(* IEC 61131-3 sources: daoli-st-library/DL_Device (part 6) *)

(* ---- FB_DL_SteamTrapMonitor.st ---- *)
(*==============================================================================
 * 组件名称 (Component)  : FB_DL_SteamTrapMonitor
 * 溯源说明 (Provenance): 道莅 clean-room 防御性实现（IEC 61131-3 纯净实现，闭源文档仅借语义，零代码行）
 * 所属子库 (Sublibrary) : DL_Device / Diagnostic
 * 当前版本 (Version)    : 1.0.0
 * 兼容性   (Platform)   : CODESYS 3.5 / TwinCAT 3 / 汇川 InoProShop / 施耐德
 *                         Machine Expert；纯 IEC 61131-3（第 3 版），仅用
 *                         Standard.library 的 TON / ABS / LIMIT / MAX
 * 组件分类 (Category)   : 功能块（FUNCTION_BLOCK）· 疏水阀堵塞/泄漏温差诊断
 * 功能一句话 (Summary)  : 用阀前/阀后温度差判断蒸汽疏水阀是正常、蒸汽泄漏（漏汽）
 *                         还是堵塞（不通），冷态停机时冻结全部故障判定。
 *
 * 本件存在的意义 (Why this unit exists)
 *   蒸汽系统节能诊断在全库零覆盖。疏水阀失效有两种相反形态：
 *   ① 漏汽（阀芯冲蚀常开）→ 阀后也被蒸汽烫热，温差变小，能耗与管网损失上升；
 *   ② 堵塞（阀芯卡死或结垢）→ 凝水积在阀前，阀前温度跌落，机组加热能力不足。
 *   两种都表现为「温差变小」，只能靠阀前温度是否达工况来区分——这就是本件
 *   判据的核心，也是它与普通温差异常报警的区别。
 *
 * 判据（公开工程判据，clean-room）
 *   正常   : fDelta >= fDeltaNormal
 *   漏汽   : fDelta <= fDeltaLeak 且 阀前温度达工况（fTin >= fTinMin）
 *   堵塞   : 阀前温度介于冷态带与工况下限之间（fTinMin × DL_COLD_RATIO <= fTin < fTinMin）
 *            且 fDelta <= fDeltaLeak
 *   冷态   : fTin < fTinMin × DL_COLD_RATIO → **工况未建立，冻结全部判定**（信息 0177）
 *   三条判据各带 tConfirm 持续确认窗，单拍越限不迁移（A5-D1 家族）。
 *   三条判据在数值上互斥（normal 要求 fDelta >= fDeltaNormal > fDeltaLeak；
 *   leak 要求 fTin >= fTinMin，blocked 要求 fTin < fTinMin），故不存在双判据
 *   同拍成立的两难情形——这是判据设计时就消除的，不靠优先级补丁。
 *
 * 冷态与堵塞的边界（规格冲突的落地方式，必须读）
 *   规格既要求「fTin < fTinMin 为工况未建立、冻结全部判定」，又要求「fTin < fTinMin
 *   （进出口均偏低、无温差）为堵塞」——同一条判据落两处。物理上二者靠「机组是否
 *   在跑」区分，本件引脚集没有机组运行信号，故用一条**相对冷态带**切分：
 *   fTinMin × DL_COLD_RATIO（0.5）以下视为停机冷态（冻结），该带与 fTinMin 之间
 *   视为「蒸汽已引入但被凝水淹没」= 堵塞特征。DL_COLD_RATIO 为件内经验常量，
 *   已在常量注释与偏离留档中声明；有运行信号的机型应把运行位并入 bEnable。
 *
 * 边界安全 (Boundary)
 *   ① fDeltaLeak >= fDeltaNormal（判据区间为空）或参数非有限 → 故障 0343、bValid = FALSE；
 *   ② 温度非有限 → 故障 0342，**保持上次判定与全部输出**（不迁移、不清状态）；
 *   ③ 冷态 → 信息 0177，冻结判定，健康投 eUnknown；
 *   ④ 落入正常带 → 信息 0176；
 *   ⑤ 健康映射集中在一处：漏汽 → eOutOfSpec（能耗越界）；堵塞 → eMaintenanceReq
 *      （需拆检）；故障 → eFailure；冷态/失能 → eUnknown；
 *   ⑥ CASE 落 ELSE 置 0344 并回 eFault；
 *   ⑦ 三条判据各用**独立 TON 实例**，绝不共用一只（R40）。
 *
 * 错误码    : 16#0003_0176 温差判据落入正常带——信息级，正常结论
 *             16#0003_0177 工况未建立（阀前温度低于冷态带），冻结判定——信息级，防误报
 *             16#0003_0342 温度输入非有限——故障级，保持上次判定
 *             16#0003_0343 判据阈值自相矛盾（fDeltaLeak >= fDeltaNormal）——故障级，bValid = FALSE
 *             16#0003_0344 状态机落 ELSE 兜底（非法状态）——故障级，回 eFault
 * 码位总账  : 16#0003_0176 用 / 16#0003_0177 用 ｜ 16#0003_0342 用 / 16#0003_0343 用 / 16#0003_0344 用
 * 状态机    : E_DL_TrapState（eIdle / eNormal / eLeak / eBlocked / eFault），CASE 含 ELSE 兜底，
 *             ELSE 置 16#0003_0344 并回 eFault；失能无条件回 eIdle
 * 采样约定  : 每任务周期调用一次；确认窗由 tConfirm 给定，不读系统时钟
 * 依赖说明  : 仅 Standard.library；健康出口引用 E_DL_Ne107Status（引用不重声明，R70③）
 * 验收向量  : V1 阀前 170 / 阀后 155（Δ15 >= 10）持续 30 s → eNormal，bNormal = TRUE，
 *                eErr = 0176，eHealth = eOk
 *             V2 阀前 165 / 阀后 162（Δ3、阀前达工况）持续 30 s → eLeak，bSteamLeak = TRUE，
 *                eHealth = eOutOfSpec
 *             V3 阀前 70 / 阀后 68（Δ2、介于冷态带 40 与 80 之间）持续 30 s → eBlocked，
 *                bBlocked = TRUE，eHealth = eMaintenanceReq（堵塞主向量）
 *             V4 阀前 30 / 阀后 28（低于冷态带 40）→ eIdle 冻结，eErr = 0177，eHealth = eUnknown
 *                （冷态防误报主向量）
 *             V5 fDeltaLeak = 12 > fDeltaNormal = 10 → 0343，bValid = FALSE，判据不成立
 *             V6 fTout = NaN → 0342，状态与输出保持上一拍（保持主向量）
 *             V7 温差在 9.9~10.1 抖动 → 单拍越限不迁移（确认窗主向量）
 * 红线自检  : 全局变量声明零使用 / 外部变量访问零使用 / 物理地址零使用 ｜ 纯 IEC 61131-3 ｜ 无除法
 *             浮点只用大小与容差比较 ｜ 无循环 ｜ 全变量双语同行注释 ｜ ENUM + CASE
 *             含 ELSE ｜ 三只 TON 在主体前部无条件刷新 ｜ 阈值常量化，无魔法数
 * 修订历史  : 2026-11-16  v1.0.0  首版入库（R22 · 批 3 · 设备诊断）
 *============================================================================*)

(*-----------------------------------------------------------------------------
 * 枚举: E_DL_TrapState（归属本功能块，同文件发布，全库唯一定义）
 * 含义: 疏水阀诊断相位。0 起步长 10。
 *-----------------------------------------------------------------------------*)
TYPE E_DL_TrapState :
(
    eIdle    := 0,     // 待机：未使能、冷态冻结或参数非法 / Idle, disabled, frozen cold state or illegal parameters
    eNormal  := 10,    // 正常：温差达到正常下限 / Normal, the temperature drop reaches the normal limit
    eLeak    := 20,    // 漏汽：温差过小且阀前已达工况 / Leaking, small drop with a live steam upstream
    eBlocked := 30,    // 堵塞：阀前温度跌落但蒸汽已引入 / Blocked, upstream cooled although steam was admitted
    eFault   := 99     // 故障：参数矛盾或非法状态 / Fault, contradictory parameters or an illegal state
);
END_TYPE

FUNCTION_BLOCK FB_DL_SteamTrapMonitor
VAR_INPUT
    fTin         : REAL;                       // 阀前温度 [degC] / upstream temperature [degC]
    fTout        : REAL;                       // 阀后温度 [degC] / downstream temperature [degC]
    fDeltaNormal : REAL := 10.0;               // 正常最小温差 [K]，须 > 0 / normal minimum temperature drop [K], must be > 0
    fDeltaLeak   : REAL := 5.0;                // 漏汽判定温差上限 [K]，须 >= 0 且 < fDeltaNormal / leak drop ceiling [K], below fDeltaNormal
    fTinMin      : REAL := 80.0;               // 蒸汽工况最低阀前温度 [degC]，须 > 0 / minimum live steam temperature [degC], must be > 0
    tConfirm     : TIME := T#30S;              // 判据确认时间 [ms] / criterion confirm time [ms]
    bEnable      : BOOL;                       // 使能 / enable
END_VAR
VAR_OUTPUT
    fDelta       : REAL;                       // 实测温差 = 阀前 − 阀后 [K] / measured temperature drop [K]
    bNormal      : BOOL;                       // 正常判定 / normal verdict
    bSteamLeak   : BOOL;                       // 漏汽判定 / steam leak verdict
    bBlocked     : BOOL;                       // 堵塞判定 / blocked verdict
    eHealth      : E_DL_Ne107Status;           // NE107 健康分级（引用唯一属主） / NE107 health status
    eErr         : UDINT;                      // 错误码，0 表示无错 / error code, 0 means no error
    bError       : BOOL;                       // 故障级标志，仅故障级错误置位 / fault-class flag, set only on fault-level codes
    bValid       : BOOL;                       // 输出可用标志 / outputs usable flag
END_VAR
VAR
    fbNormal     : TON;                        // 正常判据确认窗，段 7 无条件刷新 [ms] / normal criterion confirm window
    fbLeak       : TON;                        // 漏汽判据确认窗，段 7 无条件刷新 [ms] / leak criterion confirm window
    fbBlocked    : TON;                        // 堵塞判据确认窗，段 7 无条件刷新 [ms] / blocked criterion confirm window
    _eState      : E_DL_TrapState := E_DL_TrapState.eIdle; // 当前相位 / current phase
    _bInit       : BOOL := FALSE;              // 首扫标志，初值 FALSE 取非判定 / first-scan flag, tested negated
    _bParamBad   : BOOL;                       // 参数非法标志 / illegal parameter flag
    _bFiniteBad  : BOOL;                       // 输入非有限标志 / non-finite input flag
    _bIllegal    : BOOL;                       // 非法状态标志 / illegal state flag
    _bCold       : BOOL;                       // 冷态（工况未建立）标志 / cold state, the operating condition is not established
    _bCondNormal : BOOL;                       // 正常判据条件 / normal criterion condition
    _bCondLeak   : BOOL;                       // 漏汽判据条件 / leak criterion condition
    _bCondBlock  : BOOL;                       // 堵塞判据条件 / blocked criterion condition
    _bBrkNormal  : BOOL;                       // 正常确认计时器断输入一拍 / normal timer one-scan break
    _bBrkLeak    : BOOL;                       // 漏汽确认计时器断输入一拍 / leak timer one-scan break
    _bBrkBlock   : BOOL;                       // 堵塞确认计时器断输入一拍 / blocked timer one-scan break
    _tConfirmUse : TIME := T#30S;              // 生效确认时间 [ms]，已钳位 / effective confirm time, clamped
    _fDeltaHeld  : REAL;                       // 温差保持量 [K] / held temperature drop [K]
    _fColdLimit  : REAL := 40.0;               // 冷态带上限 [degC] = fTinMin × 冷态比 / cold band ceiling
END_VAR
VAR CONSTANT
    DL_VAL_LIM     : REAL := 1.0E6;            // 有限性判定的绝对值上限 [degC] / finiteness ceiling [degC]
    DL_DELTA_N_MN  : REAL := 0.0;              // 正常温差下限 [K]，须严格大于 / normal drop floor, strictly greater
    DL_DELTA_L_MN  : REAL := 0.0;              // 漏汽温差下限 [K] / leak drop floor [K]
    DL_TIN_MIN_MN  : REAL := 0.0;              // 工况温度下限 [degC]，须严格大于 / live steam temperature floor, strictly greater
    DL_COLD_RATIO  : REAL := 0.5;              // 冷态带相对工况下限的比例 [倍]，件内经验值 / cold band ratio, an empirical in-unit value
    DL_DELTA_MAX   : REAL := 1000.0;           // 温差合理上限 [K]，仅用于出口钳位 / sane drop ceiling [K], outlet clamping only
    DL_CONF_MAX_MS : DINT := 3600000;          // 确认时间上限 [ms]，一小时 / confirm time ceiling, one hour
    DL_TIME_ZERO   : TIME := T#0MS;            // 时间零值基准 [ms] / time zero reference
    DL_EPS         : REAL := 1.0E-6;           // 浮点比较容差 [K] / float comparison tolerance [K]
END_VAR

(*------------------------------------------------------------------------------
 * 段 1｜每拍预置（判定输出与保持量在段 9 单点写入）
 *      Per-scan presets, the verdicts are written only in segment nine
 *-----------------------------------------------------------------------------*)
eErr         := 16#0000_0000;                  // 错误码每拍重算 / error code recomputed every scan
bError       := FALSE;                         // 故障标志每拍重算 / fault flag recomputed every scan
bValid       := FALSE;                         // 可用标志每拍重算 / usable flag recomputed every scan
bNormal      := FALSE;                         // 正常判定每拍重算 / normal verdict recomputed
bSteamLeak   := FALSE;                         // 漏汽判定每拍重算 / leak verdict recomputed
bBlocked     := FALSE;                         // 堵塞判定每拍重算 / blocked verdict recomputed
_bParamBad   := FALSE;                         // 参数非法标志预清零 / parameter flag pre-cleared
_bFiniteBad  := FALSE;                         // 非有限标志预清零 / non-finite flag pre-cleared
_bIllegal    := FALSE;                         // 非法状态标志预清零 / illegal state flag pre-cleared
_bCold       := FALSE;                         // 冷态标志预清零 / cold flag pre-cleared
_bCondNormal := FALSE;                         // 正常条件预置 FALSE / normal condition preset FALSE
_bCondLeak   := FALSE;                         // 漏汽条件预置 FALSE / leak condition preset FALSE
_bCondBlock  := FALSE;                         // 堵塞条件预置 FALSE / blocked condition preset FALSE

(*------------------------------------------------------------------------------
 * 段 2｜首扫初始化（判定从待机起，不继承任何历史结论）
 *      First-scan initialisation, no historical verdict is inherited
 *-----------------------------------------------------------------------------*)
IF NOT _bInit THEN
    _eState     := E_DL_TrapState.eIdle;       // 相位待机 / phase idle
    _fDeltaHeld := 0.0;                        // 温差保持量 0 [K] / held drop zero
    _bBrkNormal := TRUE;                       // 正常确认窗从零开始 / normal window starts from zero
    _bBrkLeak   := TRUE;                       // 漏汽确认窗从零开始 / leak window starts from zero
    _bBrkBlock  := TRUE;                       // 堵塞确认窗从零开始 / blocked window starts from zero
    _bInit      := TRUE;                       // 首扫只做一次 / the first scan runs once
END_IF

(*------------------------------------------------------------------------------
 * 段 3｜参数闸门（判据区间必须非空，否则判据无意义）
 *      Parameter gate, the criteria intervals must not be empty
 *-----------------------------------------------------------------------------*)
IF (fDeltaNormal <> fDeltaNormal) OR (ABS(fDeltaNormal) > DL_VAL_LIM) OR (fDeltaNormal <= DL_DELTA_N_MN) THEN
    _bParamBad := TRUE;                        // 正常温差非法 / normal drop illegal
END_IF
IF (fDeltaLeak <> fDeltaLeak) OR (ABS(fDeltaLeak) > DL_VAL_LIM) OR (fDeltaLeak < DL_DELTA_L_MN) THEN
    _bParamBad := TRUE;                        // 漏汽温差非法 / leak drop illegal
END_IF
IF (fDeltaLeak >= fDeltaNormal) OR ((fDeltaNormal - fDeltaLeak) <= DL_EPS) THEN
    _bParamBad := TRUE;                        // 区间为空：判据自相矛盾 / empty interval, contradictory criteria
END_IF
IF (fTinMin <> fTinMin) OR (ABS(fTinMin) > DL_VAL_LIM) OR (fTinMin <= DL_TIN_MIN_MN) THEN
    _bParamBad := TRUE;                        // 工况温度非法 / live steam temperature illegal
END_IF

(*------------------------------------------------------------------------------
 * 段 4｜温度有限性（区间判据同时拦 NaN 与 ±Inf）
 *      Temperature finiteness, the interval test catches NaN and infinity
 *-----------------------------------------------------------------------------*)
IF (fTin < -DL_VAL_LIM) OR (fTin > DL_VAL_LIM) THEN
    _bFiniteBad := TRUE;                       // 阀前温度非有限 / upstream temperature non-finite
END_IF
IF (fTout < -DL_VAL_LIM) OR (fTout > DL_VAL_LIM) THEN
    _bFiniteBad := TRUE;                       // 阀后温度非有限 / downstream temperature non-finite
END_IF

(*------------------------------------------------------------------------------
 * 段 5｜温差与冷态带（冷态带由工况下限按比例导出，件内常量）
 *      Temperature drop and the cold band derived from the live steam limit
 *-----------------------------------------------------------------------------*)
IF NOT _bFiniteBad THEN
    _fDeltaHeld := fTin - fTout;               // 实测温差 [K] / measured drop
    _fColdLimit := fTinMin * DL_COLD_RATIO;    // 冷态带上限 [degC] / cold band ceiling
    _bCold      := (fTin < _fColdLimit);       // 冷态判据：明显停机 / cold test, clearly shut down
END_IF

(*------------------------------------------------------------------------------
 * 段 6｜三条判据条件（数值上互斥：由阈值关系结构性保证，不靠优先级补丁）
 *      The three criteria are mutually exclusive by construction
 *-----------------------------------------------------------------------------*)
IF (NOT _bFiniteBad) AND (NOT _bParamBad) THEN
    _bCondNormal := (_fDeltaHeld >= fDeltaNormal);                       // 正常：温差达正常下限
    _bCondLeak   := (_fDeltaHeld <= fDeltaLeak) AND (fTin >= fTinMin);   // 漏汽：温差小且阀前已达工况
    _bCondBlock  := (_fDeltaHeld <= fDeltaLeak) AND (fTin >= _fColdLimit) AND (fTin < fTinMin); // 堵塞：蒸汽已引入但阀前跌落
END_IF

(*------------------------------------------------------------------------------
 * 段 7｜三只确认计时器无条件刷新（R40：CASE 之外每拍必调，各判据各一只）
 *      Three confirm timers refreshed unconditionally, one instance per criterion
 *-----------------------------------------------------------------------------*)
_tConfirmUse := tConfirm;                      // 确认时间直取引脚 [ms] / confirm time from the pin
IF TIME_TO_DINT(_tConfirmUse) > DL_CONF_MAX_MS THEN
    _tConfirmUse := DINT_TO_TIME(DL_CONF_MAX_MS); // 超上限钳位（无专用码位，R90 不新开码） / clamped
END_IF
IF TIME_TO_DINT(_tConfirmUse) < 0 THEN
    _tConfirmUse := DL_TIME_ZERO;              // 负时间结构性不可达，兜底为 0 / structurally unreachable fallback
END_IF

fbNormal(IN := _bCondNormal AND bEnable AND (NOT _bBrkNormal), PT := _tConfirmUse); // 正常确认窗
_bBrkNormal := FALSE;                          // 断输入拍在调用后自清 / break self-cleared after the call

fbLeak(IN := _bCondLeak AND bEnable AND (NOT _bBrkLeak), PT := _tConfirmUse); // 漏汽确认窗
_bBrkLeak := FALSE;                            // 断输入拍在调用后自清 / break self-cleared

fbBlocked(IN := _bCondBlock AND bEnable AND (NOT _bBrkBlock), PT := _tConfirmUse); // 堵塞确认窗
_bBrkBlock := FALSE;                           // 断输入拍在调用后自清 / break self-cleared

(*------------------------------------------------------------------------------
 * 段 8｜相位机（非有限拍整段跳过：保持上次判定，②）
 *      Phase machine, skipped entirely on a non-finite scan to hold the last verdict
 *-----------------------------------------------------------------------------*)
IF NOT _bFiniteBad THEN
    (* 温度坏值拍整段跳过：不迁移、不清结论，保持上次判定（②），仅由码位链报 0342 *)
    (* A non-finite scan skips the whole block, the last verdict is held *)
    IF _bParamBad THEN
        _eState := E_DL_TrapState.eFault;      // 判据自相矛盾：转故障 / contradictory criteria go to fault
    ELSIF NOT bEnable THEN
        _eState := E_DL_TrapState.eIdle;       // 失能回待机 / disabled, back to idle
        _bBrkNormal := TRUE;                   // 三只确认窗全部重启 / every window restarts
        _bBrkLeak   := TRUE;                   // 漏汽窗重启 / leak window restarts
        _bBrkBlock  := TRUE;                   // 堵塞窗重启 / blocked window restarts
    ELSE
        CASE _eState OF

            E_DL_TrapState.eIdle:                  // 待机：冷态冻结，工况建立后按判据进入
                IF _bCold THEN
                    _eState := E_DL_TrapState.eIdle; // 工况未建立，冻结（0177 在段 10） / condition not established, frozen
                ELSIF fbNormal.Q THEN
                    _eState := E_DL_TrapState.eNormal; // 进正常相 / enter normal
                ELSIF fbLeak.Q THEN
                    _eState := E_DL_TrapState.eLeak;   // 进漏汽相 / enter leak
                ELSIF fbBlocked.Q THEN
                    _eState := E_DL_TrapState.eBlocked; // 进堵塞相 / enter blocked
                END_IF

            E_DL_TrapState.eNormal:                // 正常：判据迁移
                IF _bCold THEN
                    _eState := E_DL_TrapState.eIdle;   // 工况消失，回冻结 / the condition is lost, freeze
                ELSIF fbLeak.Q THEN
                    _eState := E_DL_TrapState.eLeak;   // 转漏汽 / switch to leak
                ELSIF fbBlocked.Q THEN
                    _eState := E_DL_TrapState.eBlocked; // 转堵塞 / switch to blocked
                END_IF

            E_DL_TrapState.eLeak:                  // 漏汽：判据迁移
                IF _bCold THEN
                    _eState := E_DL_TrapState.eIdle;   // 工况消失，回冻结 / freeze again
                ELSIF fbNormal.Q THEN
                    _eState := E_DL_TrapState.eNormal; // 恢复正常 / back to normal
                ELSIF fbBlocked.Q THEN
                    _eState := E_DL_TrapState.eBlocked; // 转堵塞 / switch to blocked
                END_IF

            E_DL_TrapState.eBlocked:               // 堵塞：判据迁移
                IF _bCold THEN
                    _eState := E_DL_TrapState.eIdle;   // 工况消失（彻底冷机），回冻结 / freeze again
                ELSIF fbNormal.Q THEN
                    _eState := E_DL_TrapState.eNormal; // 恢复正常 / back to normal
                ELSIF fbLeak.Q THEN
                    _eState := E_DL_TrapState.eLeak;   // 转漏汽 / switch to leak
                END_IF

            E_DL_TrapState.eFault:                 // 故障：参数恢复即回待机
                IF (NOT _bParamBad) AND (NOT _bFiniteBad) THEN
                    _eState := E_DL_TrapState.eIdle;   // 原因消失 / the cause is gone
                END_IF

            ELSE
                _bIllegal := TRUE;                 // 标记非法状态 / flag the illegal state
                _eState   := E_DL_TrapState.eFault; // 回故障态 / back to the fault state
        END_CASE
    END_IF
END_IF

(*------------------------------------------------------------------------------
 * 段 9｜出口单点写入（判定与温差唯一写入点）
 *      Single write point of the verdicts and the temperature drop
 *-----------------------------------------------------------------------------*)
fDelta := LIMIT(-DL_DELTA_MAX, _fDeltaHeld, DL_DELTA_MAX); // 温差出口钳进合理域 [K] / the drop is clamped
bNormal    := (_eState = E_DL_TrapState.eNormal);   // 正常判定出口 / normal verdict outlet
bSteamLeak := (_eState = E_DL_TrapState.eLeak);     // 漏汽判定出口 / leak verdict outlet
bBlocked   := (_eState = E_DL_TrapState.eBlocked);  // 堵塞判定出口 / blocked verdict outlet

(*------------------------------------------------------------------------------
 * 段 10｜码位优先级链与健康分级（映射集中在此，不散落实现体）
 *      Code priority chain and health grading, the mapping lives in one place
 *-----------------------------------------------------------------------------*)
IF _bIllegal THEN
    eErr   := 16#0003_0344;                    // 故障级：状态机兜底 / fault: state machine fallback
    bError := TRUE;                            // 置故障标志 / raise the fault flag
ELSIF _bParamBad THEN
    eErr   := 16#0003_0343;                    // 故障级：判据阈值自相矛盾 / fault: contradictory thresholds
    bError := TRUE;                            // 置故障标志 / raise the fault flag
ELSIF _bFiniteBad THEN
    eErr   := 16#0003_0342;                    // 故障级：温度输入非有限 / fault: non-finite temperature
    bError := TRUE;                            // 置故障标志 / raise the fault flag
ELSIF _bCold THEN
    eErr   := 16#0003_0177;                    // 信息级：工况未建立，冻结判定 / informational: condition not established
ELSIF _eState = E_DL_TrapState.eNormal THEN
    eErr   := 16#0003_0176;                    // 信息级：判据落入正常带 / informational: inside the normal band
END_IF

IF _bParamBad OR _bFiniteBad OR _bIllegal THEN
    eHealth := E_DL_Ne107Status.eFailure;      // 无判定能力：失效 / no verdict capability
ELSIF _eState = E_DL_TrapState.eLeak THEN
    eHealth := E_DL_Ne107Status.eOutOfSpec;    // 漏汽：能耗与管网越界，仍可运行 / leaking, out of specification
ELSIF _eState = E_DL_TrapState.eBlocked THEN
    eHealth := E_DL_Ne107Status.eMaintenanceReq; // 堵塞：需拆检 / blocked, maintenance required
ELSIF (_eState = E_DL_TrapState.eNormal) AND bEnable THEN
    eHealth := E_DL_Ne107Status.eOk;           // 正常 / normal
ELSE
    eHealth := E_DL_Ne107Status.eUnknown;      // 冷态或失能：无结论 / cold or disabled, no verdict
END_IF

IF bError THEN
    bValid := FALSE;                           // 故障级：输出不可用 / fault: outputs unusable
ELSIF _bCold THEN
    bValid := FALSE;                           // 冷态：判定被冻结，输出不可用 / cold: the verdict is frozen
ELSIF NOT bEnable THEN
    bValid := FALSE;                           // 失能：输出不可用 / disabled: unusable
ELSE
    bValid := TRUE;                            // 判定可用 / verdict usable
END_IF

END_FUNCTION_BLOCK

(* ---- FB_DL_StrainThermalCreepAdaptive.st ---- *)
(*
    FB_DL_StrainThermalCreepAdaptive —— 应变桥温漂与蠕变自适应补偿（含空载窗口自动重学零点）
    ------------------------------------------------------------------
    组件名    : FB_DL_StrainThermalCreepAdaptive
    分类      : DL_Device / Weighing Compensation（称重与测力补偿）
    一句话功能: 在线扣除应变桥的温漂与载荷蠕变，并在空载窗口自动重学零点，
                同时用「载荷是否真为空」判据防止把真实载荷学成漂移。
    复杂度    : C3
    版本      : v1.0.0
    开源溯源  : 无（clean-room 自研，未借鉴任何开源实现）
    平台      : 纯 IEC 61131-3（TON / R_TRIG / ABS / TIME_TO_REAL 标准转换），目标编译器
                RuSTy 1.0.8，兼容 CODESYS 3.5 / TwinCAT 3 / 汇川 InoProShop / Machine Expert；
                无 PROPERTY、无 VLA、无 FOR..DOWNTO、无 AS 类方言
    ------------------------------------------------------------------
    功能说明  : ① 温漂：fTempCorrMv = fTempCoefMvPerC × (fTempC − fRefTempC)，从原始桥压减掉；
                ② 零点：fCorrected = fRawMv − fTempCorrMv − fZeroMv，零点由空载学习维护；
                ③ 蠕变：fCreepCorrMv = fCorrected × fCreepCoefPctPerMin × 0.01 × tHoldMin，
                   方向随 fCorrected 的符号自动跟随载荷方向（负载荷得到负补偿量）；
                ④ 空载学习：bNoLoadWindow = TRUE 且持续 ≥ tLearnMinMs（TON 无条件刷新）→ 进
                   eLearn，用一阶低通（系数固定 0.05，见代理假设）把「温漂修正后、零点修正前」
                   的值学成新零点；窗口消失立即退出并冻结零点；
                ⑤ 防误学：学习期间若 |温漂修正后值| 超 fNoLoadMaxMv（载荷比 > 1）→ 判「并非空载」，
                   退出 eLearn 回 eRun 并置 bLearnRejected 单拍位；同一空载窗口内不再重试
                   （_bRejLatch 在窗口消失时清除），避免窗口内反复进出打摆；
                ⑥ 温度或原始值非有限 → eFault，且 fOutMv 保持上一次有效值（保持而非清零）。
    量纲链    : fTempCoefMvPerC [mV/°C] × (fTempC − fRefTempC) [°C] → fTempCorrMv [mV]（°C 约去）；
                fRawMv [mV] − fTempCorrMv [mV] → _fRawTemp [mV]（零点修正前）；
                _fRawTemp [mV] − fZeroMv [mV] → fCorrected [mV]（零点修正后）；
                fCorrected [mV] × fCreepCoefPctPerMin [%/min] × 0.01 [1/%] × tHoldMin [min]
                    → fCreepCorrMv [mV]（%/min × min = %，× 0.01 无因次，只剩 mV）；
                fOutMv = fCorrected [mV] − fCreepCorrMv [mV] → [mV]；
                _fLoadRatio = |_fRawTemp| [mV] ÷ _fNoLoadGuard [mV] → [-]（判载荷比与 1.0 直比）。
                全程无「温度与毫伏相加」「时间与毫伏相加」，量纲链逐段闭合。
    代理假设  : （R95 三句声明）① 代理值 = 低通系数固定 0.05，隐含标称扫描周期 10 ms，
                对应零点学习时间常数 τ ≈ 0.2 s；② 覆盖范围 = 5 ms ~ 20 ms 的周期任务
                （时间常数随之在 0.1 s ~ 0.4 s 间变化，只影响学习快慢，不影响零点收敛方向）；
                ③ 覆盖不到的区间（< 2 ms 或 > 50 ms 的任务）由现场加长 tLearnMinMs 与空载窗口
                驻留时长补偿，本件不提供自适应系数。
    交付门槛  : 本件使用 TIME_TO_REAL 标准转换做承载时长换算，须在 CODESYS / TwinCAT /
                InoProShop 三平台各编译验证一次（R64）。
    状态机    : eInit(0) --使能且输入有限且组态合法--> eRun(10)
                eRun --空载窗口持续到（tonLearn.Q）且本窗口未拒学过--> eLearn(20)
                eLearn --窗口消失--> eRun（零点冻结）；--载荷比 > 1--> eRun（拒学 + 单拍位）
                eRun/eLearn --失能--> eHold(30)（冻结保持末次有效输出与累计）
                eHold --重新使能--> eRun
                任意相 --输入非有限或组态非法--> eFault(90)
                eFault 的唯一解除路径 = bReset 上升沿（见段 8 与复位作用域声明）
    失能语义  : bEnable = FALSE → eHold，fOutMv 冻结保持末次有效值，蠕变累计与零点学习全部冻结
                （取「冻结保持」而非「降级清零」：称重输出清零会被上位当作零载荷，属伪造计量事实）。
    复位作用域: bReset 上升沿①清 _bFaultLatch / _bBadIn / _bCfgBad；②清 _fZero 与
                _fHoldBaseMin（零点与承载累计一并归零，须重新学习）；③清 _bRejLatch；
                ④迁相回 eInit；⑤不清 _fOutHold（补偿输出不因复位跳变），_bHoldValid 保留。
    防御口径  : NaN 用自反 f<>f；±Inf 用 (f−f)<>(f−f)；另设幅值域闸 ABS(f) > 1.0E30。
                除子三类：DL_ST_MS_PER_MIN = 60000.0 与 DL_ST_PCT_TO_RATIO = 0.01 为具名常量，
                结构上不可能为零；载荷比除子 _fNoLoadGuard 由 fNoLoadMaxMv 经两级下限兜底后
                才参与除法（R117 两级回退）。
                计算结果写入保持槽 _fOutHold 之前必须过非有限闸（R133），污染数据不进保持槽。
    规格偏离  : 派单把学习最短时长写作 fLearnMinMs，其实际类型为 TIME；本库规范 1.2 规定
                时间量前缀为 t，故落为 tLearnMinMs，语义不变。按 R190 归因唯一补充
                bCfgErr / bDataErr 两个诊断位，使两条故障成因各自可观测。
    码位说明  : 本件按零码位范式交付，不分配 16# 事件码；学习结果与故障一律经
                eState / bLearnRejected / bFaultOut / bCfgErr / bDataErr 组合观测。
    修订记录  : 2026-11-24 v1.0.0 首次入库（R87 批 · #3）
*)
TYPE E_DL_StrainCompState :
(
    eInit   := 0,     // 初始化：首扫或复位后，尚无可信输出 | init, no trustworthy output yet
    eRun    := 10,    // 运行：温漂 + 零点 + 蠕变三项全补偿 | running, thermal, zero and creep all compensated
    eLearn  := 20,    // 学习：空载窗口内低通重学零点，蠕变累计冻结 | learning the zero in a no-load window
    eHold   := 30,    // 保持：失能冻结末次有效输出与累计 | hold, disabled, last valid output frozen
    eFault  := 90     // 故障：输入非有限或组态非法，锁存至复位沿 | fault latched until the reset edge
);
END_TYPE

FUNCTION_BLOCK FB_DL_StrainThermalCreepAdaptive
VAR_INPUT
    bEnable             : BOOL;                   // 使能电平，TRUE = 允许补偿与学习 | enable level, TRUE = compensation and learning
    bReset              : BOOL;                   // 复位请求，上升沿生效 | reset request, rising-edge active
    fRawMv              : REAL;                   // 应变桥原始输出 [mV] | raw bridge output [mV]
    fTempC              : REAL;                   // 桥体温度 [°C] | bridge temperature [degC]
    fRefTempC           : REAL := 20.0;           // 参考温度（补偿零点温度）[°C] | reference temperature [degC]
    fTempCoefMvPerC     : REAL := 0.0;            // 温度系数 [mV/°C]，正负均合法 | temperature coefficient [mV/degC]
    fCreepCoefPctPerMin : REAL := 0.0;            // 蠕变系数 [%/min]，须非负 | creep coefficient [%/min], non-negative
    bNoLoadWindow       : BOOL;                   // 空载窗口（上位给出：工位确认为空载）| no-load window from the supervisor
    tLearnMinMs         : TIME := T#2S;           // 空载最短驻留时长，达到才允许学习 [ms] | minimum no-load dwell [ms]
    fNoLoadMaxMv        : REAL := 0.5;            // 空载带半宽，超出即判非空载 [mV] | no-load band half width [mV]
END_VAR
VAR_OUTPUT
    eState              : E_DL_StrainCompState;          // 主状态，供 HMI 使用 | main state for HMI
    fOutMv              : REAL;                   // 补偿后输出（去皮净载荷）[mV] | compensated output [mV]
    fTempCorrMv         : REAL;                   // 本拍温漂补偿量 [mV] | thermal correction this scan [mV]
    fCreepCorrMv        : REAL;                   // 本拍蠕变补偿量 [mV] | creep correction this scan [mV]
    fZeroMv             : REAL;                   // 当前生效零点 [mV] | active zero offset [mV]
    bLearnRejected      : BOOL;                   // 学习被拒事件位，单拍 | learning rejection event, single scan
    bFaultOut           : BOOL;                   // 故障汇总位 | fault aggregate
    bCfgErr             : BOOL;                   // 组态非法诊断位（归因唯一，R190）| bad-configuration flag
    bDataErr            : BOOL;                   // 数据非有限诊断位（归因唯一，R190）| non-finite data flag
END_VAR
VAR
    rtReset             : R_TRIG;                 // 复位上升沿实例，每拍无条件刷新 | reset rising-edge instance
    tonHold             : TON;                    // 承载时长分片计时，自复位，每拍无条件刷新 | load-hold slice timer, self-resetting
    tonLearn            : TON;                    // 空载窗口驻留计时，每拍无条件刷新 | no-load dwell timer
    _eState             : E_DL_StrainCompState := E_DL_StrainCompState.eInit; // 状态机内部当前态 | internal current state
    _bInit              : BOOL := TRUE;           // 首扫初始化标志，含零点与累计状态 | first-scan init flag
    _bResetLatch        : BOOL := FALSE;          // 复位沿锁存量，本拍末清除 | reset-edge latch, cleared at scan end
    _bFaultLatch        : BOOL := FALSE;          // 故障锁存位 | fault latch
    _bBadIn             : BOOL := FALSE;          // 输入非有限成因位 | non-finite input cause
    _bCfgBad            : BOOL := FALSE;          // 组态非法成因位 | bad configuration cause
    _bRejLatch          : BOOL := FALSE;          // 拒学锁存，空载窗口消失时清除 | rejection latch, cleared when the window drops
    _bHoldValid         : BOOL := FALSE;          // 保持槽已有有效值标志 | holder contains a valid value
    _bLoadNow           : BOOL := FALSE;          // 本拍存在载荷（超空载带）| load present this scan
    _fZero              : REAL := 0.0;            // 学习得到的零点 [mV] | learned zero offset [mV]
    _fTempCorr          : REAL := 0.0;            // 温漂补偿量 [mV] | thermal correction [mV]
    _fRawTemp           : REAL := 0.0;            // 温漂修正后、零点修正前的值 [mV] | thermally corrected, pre-zero [mV]
    _fCorrected         : REAL := 0.0;            // 温漂与零点均修正后的值 [mV] | fully corrected value [mV]
    _fCreepCorr         : REAL := 0.0;            // 蠕变补偿量 [mV] | creep correction [mV]
    _fOut               : REAL := 0.0;            // 本拍补偿输出 [mV] | compensated output this scan [mV]
    _fOutHold           : REAL := 0.0;            // 输出保持槽，只写已过非有限闸的值 [mV] | output holder, gated before writing [mV]
    _fNoLoadGuard       : REAL := 0.0;            // 空载带半宽的兜底值 [mV]，作除法除子 | no-load band with floor, used as divisor [mV]
    _fLoadRatio         : REAL := 0.0;            // 载荷比 [-] = |值| ÷ 空载带半宽 | load ratio, dimensionless
    _fHoldBaseMin       : REAL := 0.0;            // 已满片承载时长基值 [min] | accumulated whole-slice hold time [min]
    _fHoldMin           : REAL := 0.0;            // 参与蠕变计算的承载时长 [min] | hold time used by the creep model [min]
END_VAR
VAR CONSTANT
    DL_ST_EPS           : REAL := 1.0E-6;         // 浮点判零容差 [mV] | float zero tolerance [mV]
    DL_ST_MAG_MAX       : REAL := 1.0E30;         // 有限幅值域闸上限 [mV] | magnitude domain bound [mV]
    DL_ST_BAND_FLOOR    : REAL := 1.0E-3;         // 空载带半宽下限兜底 [mV] | no-load band floor [mV]
    DL_ST_LPF_ALPHA     : REAL := 0.05;           // 零点学习低通系数 [-]，见代理假设三句 | zero-learning low-pass coefficient
    DL_ST_MS_PER_MIN    : REAL := 60000.0;        // 毫秒与分钟换算常量 [ms/min] | milliseconds per minute
    DL_ST_PCT_TO_RATIO  : REAL := 0.01;           // 百分数转无因次常量 [1/%] | percent to ratio constant
    DL_ST_SLICE_MIN     : REAL := 60.0;           // 承载时长分片宽度 [min]（对应 TON 的 1 h 量程）| hold slice width [min]
    DL_ST_HOLD_MAX_MIN  : REAL := 1000000.0;      // 承载时长基值饱和上限 [min]，防浮点溢出 | hold-time saturation bound [min]
END_VAR

METHOD ClampToBand : REAL
(*
    把补偿量钳到 ±带宽，防止系数误配时补偿量把输出打穿。纯函数，无跨拍状态。
    Clamp a correction to a symmetric band so a mis-parameterised coefficient cannot saturate the output.
*)
VAR_INPUT
    fIn   : REAL;                                 // 待钳补偿量 [mV] | correction to clamp [mV]
    fBand : REAL;                                 // 对称带宽（已兜底为正）[mV] | symmetric band, floored positive [mV]
END_VAR
ClampToBand := fIn;                               // 直通后按两侧硬界饱和 | straight-through, saturated below
IF ClampToBand > fBand THEN
    ClampToBand := fBand;                         // 正向钳到 +带宽 [mV] | clamp to the positive band
END_IF
IF ClampToBand < (0.0 - fBand) THEN
    ClampToBand := 0.0 - fBand;                   // 负向钳到 −带宽 [mV] | clamp to the negative band
END_IF
END_METHOD

// 段 1｜输出预置与首扫初始化（含零点与累计状态，故必须有 _bInit，R310）
// segment 1, output presets and first-scan initialisation; the zero and accumulators require _bInit
fTempCorrMv := 0.0;                                // 预置温漂补偿 0 [mV] | preset zero thermal correction [mV]
fCreepCorrMv := 0.0;                               // 预置蠕变补偿 0 [mV] | preset zero creep correction [mV]
bLearnRejected := FALSE;                           // 预置无拒学事件（清零归属本段，R256）| preset no rejection event
_bBadIn := FALSE;                                  // 预置输入有限 | preset finite input
_bCfgBad := FALSE;                                 // 预置组态合法 | preset legal configuration
_bLoadNow := FALSE;                                // 预置无载荷 | preset no load
IF _bInit THEN
    _bInit := FALSE;                               // 首扫只执行一次 | runs once on the first scan
    _eState := E_DL_StrainCompState.eInit;                // 首扫状态回初相 | initialise the state
    _fZero := 0.0;                                 // 首扫零点归零 [mV]，由空载学习建立 | initial zero [mV]
    _fHoldBaseMin := 0.0;                          // 首扫承载时长归零 [min] | initial hold time [min]
    _fHoldMin := 0.0;                              // 首扫参与量归零 [min] | initial hold time for the model [min]
    _bRejLatch := FALSE;                           // 首扫清拒学锁存 | clear the rejection latch
    _bHoldValid := FALSE;                          // 首扫无有效保持值 | no valid holder value yet
END_IF

// 段 2｜非有限闸：NaN 自反 + Inf 自减 + 幅值域，逐个浮点入参枚举（R4 / R151 / R272）
// segment 2, non-finite gate over every REAL input: NaN self-reflexive, Inf by self-subtraction, magnitude bound
IF (fRawMv <> fRawMv) OR ((fRawMv - fRawMv) <> (fRawMv - fRawMv)) THEN
    _bBadIn := TRUE;                               // 原始桥压 NaN 或 ±Inf | raw bridge output NaN or infinity
END_IF
IF ABS(fRawMv) > DL_ST_MAG_MAX THEN
    _bBadIn := TRUE;                               // 原始桥压超幅值域 | raw bridge output beyond the magnitude domain
END_IF
IF (fTempC <> fTempC) OR ((fTempC - fTempC) <> (fTempC - fTempC)) THEN
    _bBadIn := TRUE;                               // 温度 NaN 或 ±Inf | temperature NaN or infinity
END_IF
IF ABS(fTempC) > DL_ST_MAG_MAX THEN
    _bBadIn := TRUE;                               // 温度超幅值域 | temperature beyond the magnitude domain
END_IF
IF (fRefTempC <> fRefTempC) OR ((fRefTempC - fRefTempC) <> (fRefTempC - fRefTempC)) THEN
    _bBadIn := TRUE;                               // 参考温度 NaN 或 ±Inf | reference temperature NaN or infinity
END_IF
IF ABS(fRefTempC) > DL_ST_MAG_MAX THEN
    _bBadIn := TRUE;                               // 参考温度超幅值域 | reference temperature beyond the magnitude domain
END_IF
IF (fTempCoefMvPerC <> fTempCoefMvPerC) OR ((fTempCoefMvPerC - fTempCoefMvPerC) <> (fTempCoefMvPerC - fTempCoefMvPerC)) THEN
    _bBadIn := TRUE;                               // 温度系数 NaN 或 ±Inf | temperature coefficient NaN or infinity
END_IF
IF ABS(fTempCoefMvPerC) > DL_ST_MAG_MAX THEN
    _bBadIn := TRUE;                               // 温度系数超幅值域 | temperature coefficient beyond the magnitude domain
END_IF
IF (fCreepCoefPctPerMin <> fCreepCoefPctPerMin) OR ((fCreepCoefPctPerMin - fCreepCoefPctPerMin) <> (fCreepCoefPctPerMin - fCreepCoefPctPerMin)) THEN
    _bBadIn := TRUE;                               // 蠕变系数 NaN 或 ±Inf | creep coefficient NaN or infinity
END_IF
IF ABS(fCreepCoefPctPerMin) > DL_ST_MAG_MAX THEN
    _bBadIn := TRUE;                               // 蠕变系数超幅值域 | creep coefficient beyond the magnitude domain
END_IF
IF (fNoLoadMaxMv <> fNoLoadMaxMv) OR ((fNoLoadMaxMv - fNoLoadMaxMv) <> (fNoLoadMaxMv - fNoLoadMaxMv)) THEN
    _bBadIn := TRUE;                               // 空载带半宽 NaN 或 ±Inf | no-load band NaN or infinity
END_IF
IF ABS(fNoLoadMaxMv) > DL_ST_MAG_MAX THEN
    _bBadIn := TRUE;                               // 空载带半宽超幅值域 | no-load band beyond the magnitude domain
END_IF

// 段 3｜组态闸与两级兜底：空载带半宽作除法除子，先兜底；蠕变系数须非负；学习时长须非负
// segment 3, configuration gate and two-stage fallback; the band is a divisor and the creep coefficient must be non-negative
_fNoLoadGuard := fNoLoadMaxMv;                     // 取配置空载带半宽 [mV] | take the configured band [mV]
IF _fNoLoadGuard < DL_ST_BAND_FLOOR THEN
    _fNoLoadGuard := DL_ST_BAND_FLOOR;             // 一级兜底：钳到定义域下限 [mV] | stage-one clamp to the floor [mV]
END_IF
IF fCreepCoefPctPerMin < 0.0 THEN
    _bCfgBad := TRUE;                              // 蠕变系数为负：方向无物理意义，判组态非法 | negative creep coefficient is illegal
END_IF
IF tLearnMinMs < T#0S THEN
    _bCfgBad := TRUE;                              // 学习时长非法（TIME 负值）：判组态非法 | negative learning time is illegal
END_IF
IF fNoLoadMaxMv <= DL_ST_EPS THEN
    _bCfgBad := TRUE;                              // 空载带为零或负：空载判据无法成立，判组态非法 | degenerate band is illegal
END_IF

// 段 4｜温漂修正与零点修正（双闸均通过才计算，避免污染下游全部判据）
// segment 4, thermal and zero correction; computed only when both gates pass, so no polluted value flows downstream
IF (NOT _bBadIn) AND (NOT _bCfgBad) THEN
    _fTempCorr := fTempCoefMvPerC * (fTempC - fRefTempC); // 温漂补偿量 [mV] = [mV/°C] × [°C] | thermal correction [mV]
    _fRawTemp := fRawMv - _fTempCorr;              // 温漂修正后、零点修正前 [mV] | thermally corrected, pre-zero [mV]
    _fCorrected := _fRawTemp - _fZero;             // 零点修正后 [mV] | zero-corrected [mV]
    _fLoadRatio := ABS(_fRawTemp) / _fNoLoadGuard; // 载荷比 [-] = [mV] ÷ [mV]，除子已兜底非零 | guarded division
    IF _fLoadRatio > 1.0 THEN
        _bLoadNow := TRUE;                         // 超空载带：判定存在载荷 | beyond the band, load present
    END_IF
ELSE
    _fTempCorr := 0.0;                             // 闸门未过：本拍补偿量置 0，输出走保持 | gates failed, correction zeroed
    _fCorrected := 0.0;                            // 闸门未过：修正值为 0 且不写入保持槽 | corrected value zeroed, not stored
    _fLoadRatio := 0.0;                            // 闸门未过：载荷比置 0 | load ratio zeroed
END_IF

// 段 5｜定时器与沿实例无条件周期刷新（R7）；承载计时自复位（R188）
// segment 5, timers and edge instances refreshed unconditionally; the hold-slice timer is self-resetting
rtReset(CLK := bReset);
tonHold(IN := (NOT tonHold.Q) AND bEnable AND (NOT _bFaultLatch) AND _bLoadNow AND (_eState <> E_DL_StrainCompState.eLearn), PT := T#1H);
tonLearn(IN := bEnable AND bNoLoadWindow AND (NOT _bFaultLatch) AND (NOT _bRejLatch), PT := tLearnMinMs);
IF rtReset.Q THEN
    _bResetLatch := TRUE;                          // 复位沿存锁存量，段 8 统一消费 | store the reset edge, consumed in segment 8
END_IF

// 段 6｜承载时长累计：分片到时分片基值 +1，未满片的零头按 ET 折分钟（边界拍去重，R45②）
// segment 6, hold-time accumulation; whole slices are added to the base, the remainder comes from ET without double counting
IF tonHold.Q THEN
    _fHoldBaseMin := _fHoldBaseMin + DL_ST_SLICE_MIN; // 满一个分片：基值加 60 [min] | one slice completed, add 60 min
    IF _fHoldBaseMin > DL_ST_HOLD_MAX_MIN THEN
        _fHoldBaseMin := DL_ST_HOLD_MAX_MIN;        // 饱和，防浮点溢出 | saturate to avoid float overflow
    END_IF
    _fHoldMin := _fHoldBaseMin;                    // 到时分片已计入基值，ET 不再重复折算 | the slice is already in the base
ELSE
    _fHoldMin := _fHoldBaseMin + TIME_TO_REAL(tonHold.ET) / DL_ST_MS_PER_MIN; // 基值 + 零头 [min]，除子为常量 | base plus remainder [min]
END_IF

// 段 7｜空载窗口消失即解除拒学锁存（唯一清除边；否则同一窗口内永久拒学）
// segment 7, dropping the no-load window clears the rejection latch, the only release edge for that latch
IF NOT bNoLoadWindow THEN
    _bRejLatch := FALSE;                           // 窗口消失 → 下一窗口可重试学习 | window dropped, the next window may retry
END_IF

// 段 8｜复位沿与故障锁存（复位先执行，保证本拍新故障不被抹除，R275）
// segment 8, reset edge and fault latches; reset runs first so a same-scan fault survives
IF _bResetLatch THEN
    _bFaultLatch := FALSE;                         // 清故障锁存 | clear the fault latch
    _bBadIn := FALSE;                              // 清数据非有限成因位 | clear the non-finite cause
    _bCfgBad := FALSE;                             // 清组态非法成因位（下一拍按新参数重判）| clear the configuration cause
    _fZero := 0.0;                                 // 零点归零 [mV]，须重新学习 | zero cleared, must be re-learned
    _fHoldBaseMin := 0.0;                          // 承载累计归零 [min] | hold-time base cleared
    _fHoldMin := 0.0;                              // 参与量归零 [min] | hold time for the model cleared
    _bRejLatch := FALSE;                           // 清拒学锁存 | clear the rejection latch
    _eState := E_DL_StrainCompState.eInit;                // 迁相回初相 | return to the init phase
END_IF
IF _bBadIn AND (NOT _bFaultLatch) THEN
    _bFaultLatch := TRUE;                          // 锁存数据非有限（独立成因）| latch the non-finite cause
    _eState := E_DL_StrainCompState.eFault;               // 与锁存同拍迁相（R258）| migrate in the same scan
END_IF
IF _bCfgBad AND (NOT _bFaultLatch) THEN
    _bFaultLatch := TRUE;                          // 锁存组态非法（独立成因）| latch the configuration cause
    _eState := E_DL_StrainCompState.eFault;               // 与锁存同拍迁相（R258）| migrate in the same scan
END_IF

// 段 9｜主状态机：ENUM + CASE + ELSE 兜底（R6）
// segment 9, main state machine with ENUM + CASE + ELSE fallback
CASE _eState OF
E_DL_StrainCompState.eInit:
    // 拍 N 进入：首扫或复位沿；本拍行为：不做补偿写入，保持槽尚未建立；
    // 拍 N+1 转出：使能且输入有限且组态合法 → eRun
    // entered on the first scan or the reset edge; no compensation is written yet because the holder is empty;
    // exits to eRun once enabled with finite inputs and a legal configuration
    IF bEnable AND (NOT _bBadIn) AND (NOT _bCfgBad) THEN
        _eState := E_DL_StrainCompState.eRun;
    END_IF

E_DL_StrainCompState.eRun:
    IF NOT bEnable THEN
        _eState := E_DL_StrainCompState.eHold;            // 失能 → 保持相 | disable falls into hold
    ELSIF bNoLoadWindow AND tonLearn.Q THEN
        _eState := E_DL_StrainCompState.eLearn;           // 空载窗口驻留到且本窗口未拒学 → 进学习 | dwell elapsed, enter learning
    END_IF

E_DL_StrainCompState.eLearn:
    // 学习：低通把「温漂修正后、零点修正前」的值学成零点；该值不含零点自身，故不会自激
    // learning: the low-pass tracks the thermally corrected pre-zero value, which excludes the zero itself
    IF NOT bEnable THEN
        _eState := E_DL_StrainCompState.eHold;            // 失能 → 保持相（零点冻结）| disable falls into hold, the zero is frozen
    ELSIF NOT bNoLoadWindow THEN
        _eState := E_DL_StrainCompState.eRun;             // 窗口消失 → 退出并冻结零点 | the window dropped, freeze the zero
    ELSIF _fLoadRatio > 1.0 THEN
        bLearnRejected := TRUE;                    // 拒学事件，单拍（清零归属段 1）| rejection event, single scan
        _bRejLatch := TRUE;                        // 本窗口内不再重试 | no retry inside this window
        _eState := E_DL_StrainCompState.eRun;             // 回运行相，零点保持旧值 | back to run with the previous zero
    ELSE
        _fZero := _fZero + DL_ST_LPF_ALPHA * (_fRawTemp - _fZero); // 零点一阶低通 [mV] | first-order zero tracking [mV]
    END_IF

E_DL_StrainCompState.eHold:
    // 保持：不学习、不累计、不更新保持槽；fOutMv 由 _fOutHold 回放（冻结保持，见头注释失能语义）
    // hold: no learning, no accumulation and no holder update; the output replays the frozen holder
    IF bEnable AND (NOT _bFaultLatch) THEN
        _eState := E_DL_StrainCompState.eRun;             // 重新使能 → 回运行相 | re-enabled, back to run
    END_IF

E_DL_StrainCompState.eFault:
    // 驻留语义：本相只能由段 8 的复位沿迁出（唯一解除路径）；输出保持末次有效值
    // dwell semantics: left only through the reset edge in segment 8; the output keeps the last valid value

ELSE
    // 非法枚举值（越界或未定义成员）：不猜，置故障并回故障相
    // illegal enumerator: no guessing, latch a fault and return to the fault phase
    _bFaultLatch := TRUE;
    _eState := E_DL_StrainCompState.eFault;
END_CASE;

// 段 10｜蠕变补偿与保持槽写入（写入前过非有限闸，R133；组态闸与数据闸均通过才写）
// segment 10, creep correction and holder write; the value is gated before it enters the holder
IF (NOT _bBadIn) AND (NOT _bCfgBad) AND (NOT _bFaultLatch) THEN
    _fCreepCorr := _fCorrected * fCreepCoefPctPerMin * DL_ST_PCT_TO_RATIO * _fHoldMin; // 蠕变补偿 [mV]，符号随载荷 | creep correction [mV]
    _fCreepCorr := ClampToBand(_fCreepCorr, ABS(_fCorrected)); // 钳到 ±|当前载荷|，系数误配时不得把输出打穿 | clamp to the load magnitude
    _fOut := _fCorrected - _fCreepCorr;            // 补偿输出 [mV] = [mV] − [mV] | compensated output [mV]
    IF (_fOut <> _fOut) OR ((_fOut - _fOut) <> (_fOut - _fOut)) THEN
        _bBadIn := TRUE;                           // 输出侧兜底：结果非有限则拒收并置数据成因位 | result non-finite, reject and flag
        _bFaultLatch := TRUE;                      // 同拍锁存故障，保证 bFaultOut 与 eFault 语义一致（R256 三件套）| latch in the same scan
        _eState := E_DL_StrainCompState.eFault;           // 同拍迁相（R256 三件套之一）| migrate in the same scan
    ELSE
        IF (_eState = E_DL_StrainCompState.eRun) OR (_eState = E_DL_StrainCompState.eLearn) THEN
            _fOutHold := _fOut;                    // 只有已证明有限的值才进保持槽 | only a proven finite value enters the holder
            _bHoldValid := TRUE;                   // 保持槽已建立 | holder established
        END_IF
        // 保持相、初相与故障相不更新保持槽：失能即冻结末次有效值（头注释已声明「冻结保持」，R191）
        // the hold, init and fault phases never update the holder, which implements the declared freeze semantics
    END_IF
ELSE
    _fCreepCorr := 0.0;                            // 闸门未过：本拍蠕变补偿置 0，输出走保持 | gates failed, correction zeroed
END_IF

// 段 11｜出口单点映射（保持槽回放，非有限污染不会外泄）
// segment 11, single-point output mapping; the holder is replayed so no polluted value leaks out
eState := _eState;                                 // 状态映射 | state mapping
fTempCorrMv := _fTempCorr;                         // 温漂补偿量映射 [mV] | thermal correction mapping [mV]
fCreepCorrMv := _fCreepCorr;                       // 蠕变补偿量映射 [mV] | creep correction mapping [mV]
fZeroMv := _fZero;                                 // 生效零点映射 [mV] | active zero mapping [mV]
IF _bHoldValid THEN
    fOutMv := _fOutHold;                           // 有有效历史值：冻结保持末次有效输出 [mV] | replay the last valid output [mV]
ELSE
    fOutMv := 0.0;                                 // 从未建立有效值：输出哨兵零点，不伪造读数 [mV] | sentinel zero, never a fake reading
END_IF
bFaultOut := _bFaultLatch;                         // 故障锁存回放 | replay the fault latch
bCfgErr := _bCfgBad;                               // 组态非法诊断位 | bad-configuration diagnostic
bDataErr := _bBadIn;                               // 数据非有限诊断位 | non-finite data diagnostic

// 段 12｜本拍消费量收尾（仅清沿锁存；不触碰任何锁存位与 CASE 内写入量）
// segment 12, end-of-scan cleanup; only the edge latch is cleared
_bResetLatch := FALSE;
END_FUNCTION_BLOCK

(* ---- FB_DL_TankBlanketPrCtrl.st ---- *)
(*==============================================================================
 * 组件名称 (Component)  : FB_DL_TankBlanketPrCtrl
 * 所属子库 (Sublibrary) : DL_Device
 * 当前版本 (Version)    : 1.0.0
 * 兼容性   (Platform)   : CODESYS 3.5+ / TwinCAT 3 / 汇川 InoProShop / 施耐德 Machine Expert
 *                         仅依赖 Standard.library（TON / R_TRIG），零厂商私有库
 * 功能描述 (Function)   : 储罐氮封压差监测联动。
 *                         两只压力变送器（A/B）冗余采集氮封压差，按"双表一致 → 取均值；双表偏离超限 →
 *                         锁存传感器偏离故障并退化为**取低值**（保守侧：宁可早开补气阀，不可迟开）"
 *                         的判据链给出唯一可信压差，再驱动氮封补气阀与超压排放阀。
 *                         三条固化纪律：
 *                           ① **双表冗余判据（复用 RedundantSwitch 语义）**：本件不实例化
 *                              `FB_DL_RedundantSwitch`（R47 批次零文件级依赖），复用其三条语义——
 *                              偏差闸、退化取低值、偏离故障锁存；
 *                           ② **低压联锁**：可信压差低于低压门槛并经 tLowConf 确认后锁存 bLowInterlock，
 *                              补气阀保持开启直到压差回升到门槛 + 迟滞（迟滞防抖，不靠时间滤）；
 *                           ③ **阀输出限幅**：模拟阀位指令钳在 [fOpenMinPct, 100]，BOOL 阀位与之同源
 *                              （名实双出口，R191），禁"模拟量说开、BOOL 说关"。
 *                         验收向量：
 *                           ① 表 A=3.0 kPa、表 B=3.2 kPa、偏差限 0.5 → 一致，取均值 3.1 kPa
 *                           ② 表 A=3.0 kPa、表 B=5.0 kPa → 偏离 2.0 > 0.5，锁存偏离，取低值 3.0 kPa
 *                           ③ 低压门槛 2.0 kPa、迟滞 0.2、可信压差 1.8 且持续 tLowConf → 锁存低压联锁
 *                           ④ 压差回升到 2.25 kPa → 高于 2.0+0.2，补气阀关断、联锁解除（非锁存件复位前）
 * 接口     (Interface)  : 入 bEnable 使能、fPrRawA / fPrRawB 双表原始值、fSpanKpa 量程标定、
 *                         fDevMaxKpa 双表偏差限、fPrLowKpa 低压门槛、fPrHighKpa 超压门槛、
 *                         fHystKpa 迟滞半宽、tLowConf 低压确认时长、bReset 复位沿；
 *                         出 fPrSelected 可信压差、fPrDev 双表偏差、bMakeupValve 补气阀位、
 *                         fValveCmdPct 补气阀位指令、bVentValve 排放阀位、bLowInterlock 低压联锁锁存、
 *                         bSensorDev 双表偏离锁存、eState 相、eCause 成因、bError 故障标志。
 * 边界     (Boundary)   : ① **属主边界（写死）：本件只做"压差判据 + 阀位指令"，不驱动电磁阀线圈、
 *                         不做阀门回讯确认**（属阀件 / IO 映射层）；② **标定除零闸**：fSpanKpa ≤ 0
 *                         或非有限 → 锁存 eCfgIllegal（零量程会把任何原始值放大成无穷，R179）；
 *                         ③ **门槛单调闸**：fPrLow < fPrHigh 且 fHyst ≥ 0 且 fHyst < 门槛差的一半；
 *                         ④ **退化取低值**：双表偏离时选 min(A,B)，安全侧赋值只取"已证明可用的局部工作值"
 *                         或常量，绝不取被判非法的脚值（R127）；
 *                         ⑤ **确认 TON 冻结**：tonLowConf 的 IN 串 (NOT _bFault)，故障期不累计，
 *                         复位同拍不会立即重锁（R252）；TON 段 0 无条件调用；
 *                         ⑥ **锁存解除式**：bSensorDev 与 bLowInterlock 的解除各有独立路径——
 *                         bSensorDev 由 bReset 沿解除（需人工确认传感器）；bLowInterlock 由
 *                         "压差回升过门槛 + 迟滞"自动解除，两条都写死并自证可满足；
 *                         ⑦ 非有限样本 → 该路作废（当拍不参与均值），双路皆废 → 当拍不判、bValid=FALSE；
 *                         ⑧ 零全局耦合、零物理地址。
 * 分工声明 (Scope)      : 本件只管"氮封压差判据与阀位指令"。不接管：储罐液位控制
 *                         （属 FB_DL_TankLevelCtrl 族）、氮气纯度分析（属气体分析件）、
 *                         阀门故障诊断（属阀件）。
 * 来源标签 (Source Tag) : ROADMAP 空勾真缺口 P2（氮封压差联动，自研 clean-room）
 * 码表     (Codes)      : 本件不占用任何全局数字码位（零码位范式 R297）；诊断由 BOOL + ENUM 出口承担。
 * 红线自检 (Redline)    : R1 ✓ 零 GVL/VAR_EXTERNAL ｜ R2 ✓ 零 %I/%Q/%M ｜ R3 ✓ 纯 IEC 61131-3
 *                         R4 ✓ 零量程闸 + 门槛单调闸 + 阀位限幅 + 非有限闸 ｜ R5 ✓ 声明逐行同行双语注释
 *                         R6 ✓ ENUM+CASE 含 ELSE 兜底 ｜ R7 ✓ TON/R_TRIG 段 0 无条件刷新
 * 修订历史 (Revision)   : 2026-11-19  v1.0.0  R47 首版（批次 2 · 序号 9）
 *==============================================================================*)

TYPE E_DL_TbpState :
(
    eIdle    := 0,    // 待机相（未使能，阀位全关） / Idle, disabled, valves closed
    eMonitor := 10,   // 监测相（判据与阀位联动） / Monitoring, judgement and valve interlock
    eFault   := 90    // 故障相（等复位，阀位全关） / Fault, valves closed, awaiting reset
);
END_TYPE

TYPE E_DL_TbpCause :
(
    eNone      := 0,   // 无异常 / No anomaly
    eCfgIllegal:= 1,   // 组态非法（量程/门槛/迟滞越域） / Illegal configuration
    eSensorDev := 2,   // 双表偏离超限（锁存，取低值退化） / Transmitter deviation, latched, low value used
    eLowPr     := 3,   // 氮封低压联锁（锁存，等压差回升） / Blanket low pressure interlock, latched
    eBothBad   := 4,   // 双表皆非有限（当拍不判） / Both transmitters non-finite
    ePhaseBad  := 5    // 非法相位兜底 / Illegal phase fallback
);
END_TYPE

FUNCTION_BLOCK FB_DL_TankBlanketPrCtrl
VAR_INPUT
    bEnable    : BOOL := FALSE;      // 使能（FALSE 时阀位全关） [-] / Enable, valves closed when FALSE
    fPrRawA    : LREAL := 0.0;       // A 表原始值（按量程标定解释） [raw] / Transmitter A raw value
    fPrRawB    : LREAL := 0.0;       // B 表原始值（按量程标定解释） [raw] / Transmitter B raw value
    fSpanKpa   : LREAL := 10.0;      // 量程标定（原始值 → kPa 的比例），域 > 0 [kPa/raw] / Span calibration, > 0
    fDevMaxKpa : LREAL := 0.5;       // 双表偏差限，域 > 0 [kPa] / Transmitter deviation limit, > 0
    fPrLowKpa  : LREAL := 2.0;       // 低压联锁门槛 [kPa] / Low-pressure interlock threshold
    fPrHighKpa : LREAL := 6.0;       // 超压排放门槛，域 > 低压门槛 [kPa] / Over-pressure vent threshold
    fHystKpa   : LREAL := 0.2;       // 迟滞半宽，域 ≥ 0 [kPa] / Hysteresis half-width, >= 0
    tLowConf   : TIME := T#2S;       // 低压确认时长，域 > T#0S [ms] / Low-pressure confirmation time, > T#0S
    bReset     : BOOL := FALSE;      // 复位沿（清双表偏离锁存） [-] / Reset edge, clears the deviation latch
END_VAR
VAR_OUTPUT
    fPrSelected  : LREAL := 0.0;                          // 可信压差 [kPa] / Trusted blanket pressure [kPa]
    fPrDev       : LREAL := 0.0;                          // 双表偏差绝对值 [kPa] / Absolute transmitter deviation [kPa]
    bMakeupValve : BOOL := FALSE;                         // 补气阀位 [-] / Make-up valve position
    fValveCmdPct : LREAL := 0.0;                          // 补气阀位指令，钳 0..100 [%] / Make-up valve command, clamped 0..100
    bVentValve   : BOOL := FALSE;                         // 超压排放阀位 [-] / Vent valve position
    bLowInterlock: BOOL := FALSE;                         // 低压联锁锁存 [-] / Low-pressure interlock, latched
    bSensorDev   : BOOL := FALSE;                         // 双表偏离锁存 [-] / Transmitter deviation, latched
    bValid       : BOOL := FALSE;                         // 判据有效（至少一路有限） [-] / Judgement valid
    eState       : E_DL_TbpState := E_DL_TbpState.eIdle;  // 相出口 [-] / Phase outlet
    eCause       : E_DL_TbpCause := E_DL_TbpCause.eNone;  // 成因出口（R190 归因唯一） [-] / Cause outlet
    bError       : BOOL := FALSE;                         // 故障标志（组态级或双表皆废） [-] / Error flag
END_VAR
VAR
    _eState    : E_DL_TbpState := E_DL_TbpState.eIdle;    // 内部相（CASE 唯一写入目标） / Internal phase
    _eCause    : E_DL_TbpCause := E_DL_TbpCause.eNone;    // 成因锁存量 / Latched cause
    _bFault    : BOOL := FALSE;                           // 故障锁存位（组态级） / Latched configuration fault
    _bDevLatch : BOOL := FALSE;                           // 双表偏离锁存位 / Latched deviation bit
    _bLowLatch : BOOL := FALSE;                           // 低压联锁锁存位 / Latched low-pressure bit
    _fA        : LREAL := 0.0;                            // A 表换算后压差 [kPa] / Transmitter A converted value
    _fB        : LREAL := 0.0;                            // B 表换算后压差 [kPa] / Transmitter B converted value
    _bAOk      : BOOL := FALSE;                           // A 表可用标志 / Transmitter A usable
    _bBOk      : BOOL := FALSE;                           // B 表可用标志 / Transmitter B usable
    _fSel      : LREAL := 0.0;                            // 可信压差工作值 [kPa] / Trusted pressure working value
    _fDev      : LREAL := 0.0;                            // 偏差工作值 [kPa] / Deviation working value
    _fPct      : LREAL := 0.0;                            // 阀位指令工作值 [%] / Valve command working value
    _bMakeup   : BOOL := FALSE;                           // 补气阀内部位（迟滞保持量） / Internal make-up valve bit
    _bVent     : BOOL := FALSE;                           // 排放阀内部位（迟滞保持量） / Internal vent valve bit
    _bCfgBad   : BOOL := FALSE;                           // 组态非法当拍量 / Illegal configuration this scan
    tonLowConf : TON;                                     // 低压确认实例，段 0 无条件调用 / Low-pressure confirmation instance
    rtReset    : R_TRIG;                                  // 复位沿实例，段 0 无条件调用 / Reset edge instance
END_VAR
VAR CONSTANT
    DL_TBP_PCT_MAX  : LREAL := 100.0;     // 阀位指令上限 [%] / Valve command upper bound [%]
    DL_TBP_PCT_MIN  : LREAL := 0.0;       // 阀位指令下限 [%] / Valve command lower bound [%]
    DL_TBP_EPS      : LREAL := 1.0E-9;    // 浮点判等容差 [kPa] / Equality tolerance [kPa]
END_VAR

(* —— 段 0：组态闸 + TON 与沿无条件周期刷新（R228A；IN 串故障否决，R252） —— *)
_bCfgBad := (fSpanKpa <= 0.0) OR (fSpanKpa <> fSpanKpa)                       // 量程须为正且有限 / Span positive and finite
         OR (fDevMaxKpa <= 0.0) OR (fDevMaxKpa <> fDevMaxKpa)                 // 偏差限须为正且有限 / Deviation limit positive
         OR (NOT (fPrLowKpa < fPrHighKpa))                                    // 门槛须满足低压 < 超压 / Low threshold below high threshold
         OR (fHystKpa < 0.0) OR (fHystKpa > ((fPrHighKpa - fPrLowKpa) / 2.0)) // 迟滞须非负且小于门槛差半宽 / Hysteresis within the band
         OR (tLowConf <= T#0S);                                               // 确认时长须为正 / Confirmation time positive
rtReset(CLK := bReset);                                                       // 复位沿 / Reset edge
tonLowConf(IN := (_eState = E_DL_TbpState.eMonitor) AND (NOT _bFault), PT := tLowConf);   // 低压确认（监测相派生） / Low-pressure confirmation

(* —— 段 1：单拍/输出量预置（锁存量 _eCause/_bFault/_bDevLatch/_bLowLatch/_bMakeup/_bVent 不入清单，R107） —— *)
fPrSelected := 0.0;                                          // 可信压差预置 / Trusted pressure preset
fPrDev      := 0.0;                                          // 偏差预置 / Deviation preset
fValveCmdPct:= 0.0;                                          // 阀位指令预置 / Valve command preset
bMakeupValve:= FALSE;                                        // 补气阀预置 / Make-up valve preset
bVentValve  := FALSE;                                        // 排放阀预置 / Vent valve preset
bValid      := FALSE;                                        // 有效位预置 / Validity preset
bError      := FALSE;                                        // 故障标志预清（R45 配对） / Error preset
_fSel       := 0.0;                                          // 可信压差工作值预置 / Working value preset
_fDev       := 0.0;                                          // 偏差工作值预置 / Deviation working value preset
_fPct       := DL_TBP_PCT_MIN;                               // 阀位工作值预置为下限 / Command working value at the lower bound

(* —— 段 2：组态闸（非法即锁存，阀位全关） —— *)
IF _bCfgBad THEN
    _eCause := E_DL_TbpCause.eCfgIllegal;                    // 归因：组态非法 / Cause: illegal configuration
    _bFault := TRUE;                                         // 锁存 / Latch
    _eState := E_DL_TbpState.eFault;                         // 入故障相 / Enter fault phase
END_IF

(* —— 段 3：迁出链（bReset 清组态故障与双表偏离锁存；低压联锁不走复位，走压差回升） —— *)
IF rtReset.Q THEN
    _bFault    := FALSE;                                     // 清组态故障锁存 / Clear the configuration fault latch
    _bDevLatch := FALSE;                                     // 清双表偏离锁存（需人工确认后复位） / Clear the deviation latch
    _eCause    := E_DL_TbpCause.eNone;                       // 清成因 / Clear cause
    _eState    := E_DL_TbpState.eIdle;                       // 回待机相 / Back to idle
END_IF

(* —— 段 4：相迁移（使能驱动；故障相由段 3 迁出） —— *)
CASE _eState OF

E_DL_TbpState.eIdle:
    IF bEnable THEN
        _eState := E_DL_TbpState.eMonitor;                   // 使能即进监测相 / Enable enters monitoring
    END_IF

E_DL_TbpState.eMonitor:
    IF NOT bEnable THEN
        _eState := E_DL_TbpState.eIdle;                      // 失能回待机相（阀位在出口强制全关） / Disable returns to idle
    END_IF

E_DL_TbpState.eFault:
    ;                                                        // 故障相：由段 3 复位沿迁出 / Exit handled by the reset edge

ELSE
    _eCause := E_DL_TbpCause.ePhaseBad;                      // 归因：非法相位 / Cause: illegal phase
    _bFault := TRUE;                                         // 锁存 / Latch
    _eState := E_DL_TbpState.eFault;                         // 强拉故障相 / Force fault phase

END_CASE

(* —— 段 5：双表换算（原始值 × 量程比例；非有限路作废，双废当拍不判） —— *)
IF (_eState = E_DL_TbpState.eMonitor) AND (NOT _bCfgBad) THEN
    _bAOk := NOT ((fPrRawA <> fPrRawA) OR ((fPrRawA - fPrRawA) <> (fPrRawA - fPrRawA)));   // A 路有限 / A finite
    _bBOk := NOT ((fPrRawB <> fPrRawB) OR ((fPrRawB - fPrRawB) <> (fPrRawB - fPrRawB)));   // B 路有限 / B finite
    IF _bAOk THEN
        _fA := fPrRawA * fSpanKpa;                           // A 表换算为 kPa / Convert A to kPa
    END_IF
    IF _bBOk THEN
        _fB := fPrRawB * fSpanKpa;                           // B 表换算为 kPa / Convert B to kPa
    END_IF

    IF (NOT _bAOk) AND (NOT _bBOk) THEN
        _eCause := E_DL_TbpCause.eBothBad;                   // 归因：双表皆废（当拍不判，不锁存） / Cause: both transmitters unusable
    ELSIF (NOT _bBOk) THEN
        _fSel := _fA;                                        // 仅 A 可用：取 A（并记偏离锁存外的降级） / Only A usable
        _fDev := 0.0;                                        // 无对照：偏差按 0 报 / No reference, deviation reported as 0
        bValid := TRUE;
    ELSIF (NOT _bAOk) THEN
        _fSel := _fB;                                        // 仅 B 可用：取 B / Only B usable
        _fDev := 0.0;                                        // 无对照：偏差按 0 报 / No reference
        bValid := TRUE;
    ELSE
        _fDev := ABS(_fA - _fB);                             // 双表偏差绝对值 / Absolute deviation
        IF _fDev > fDevMaxKpa THEN
            _bDevLatch := TRUE;                              // 偏离超限：锁存 / Deviation beyond the limit: latch
            _eCause := E_DL_TbpCause.eSensorDev;             // 归因：双表偏离 / Cause: transmitter deviation
            IF _fA < _fB THEN
                _fSel := _fA;                                // 退化取低值（保守侧） / Degrade to the lower reading
            ELSE
                _fSel := _fB;                                // 退化取低值（保守侧） / Degrade to the lower reading
            END_IF
        ELSE
            _fSel := (_fA + _fB) / 2.0;                      // 双表一致：取均值 / Consistent, use the mean
        END_IF
        bValid := TRUE;
    END_IF

    (* —— 段 6：低压联锁（门槛 + 确认时长；回升过"门槛 + 迟滞"自动解除） —— *)
    IF bValid THEN
        IF (_fSel < fPrLowKpa) AND tonLowConf.Q THEN
            _bLowLatch := TRUE;                              // 低压确认到位：锁存联锁 / Confirm and latch the interlock
            _eCause := E_DL_TbpCause.eLowPr;                 // 归因：氮封低压 / Cause: blanket low pressure
        ELSIF _fSel > (fPrLowKpa + fHystKpa) THEN
            _bLowLatch := FALSE;                             // 回升过门槛 + 迟滞：自动解除 / Recovery clears the interlock
        END_IF

        (* —— 段 7：阀位联动（补气阀：低压或联锁 → 开；超压 → 关；其余按迟滞保持） —— *)
        IF _bLowLatch OR (_fSel < (fPrLowKpa - fHystKpa)) THEN
            _bMakeup := TRUE;                                // 低压侧：补气阀开 / Low side: open the make-up valve
        ELSIF _fSel > (fPrLowKpa + fHystKpa) THEN
            _bMakeup := FALSE;                               // 回升：补气阀关 / Recovered: close the make-up valve
        END_IF

        IF _fSel > fPrHighKpa THEN
            _bVent := TRUE;                                  // 超压：排放阀开 / Over-pressure: open the vent valve
        ELSIF _fSel < (fPrHighKpa - fHystKpa) THEN
            _bVent := FALSE;                                 // 回落：排放阀关 / Below the hysteresis: close the vent
        END_IF

        (* —— 段 8：阀位指令限幅（开则满开、关则零，指令与 BOOL 同源） —— *)
        IF _bMakeup THEN
            _fPct := DL_TBP_PCT_MAX;                         // 开阀指令 100 % / Open command
        ELSE
            _fPct := DL_TBP_PCT_MIN;                         // 关阀指令 0 % / Close command
        END_IF
        IF _fPct > DL_TBP_PCT_MAX THEN
            _fPct := DL_TBP_PCT_MAX;                         // 上钳 / Clamp high
        ELSIF _fPct < DL_TBP_PCT_MIN THEN
            _fPct := DL_TBP_PCT_MIN;                         // 下钳 / Clamp low
        END_IF
    ELSE
        _bMakeup := FALSE;                                   // 判据无效：补气阀保守关（不猜方向） / Invalid: close conservatively
        _bVent   := FALSE;                                   // 判据无效：排放阀关 / Invalid: vent closed
        _fPct    := DL_TBP_PCT_MIN;                           // 指令归零 / Command zeroed
    END_IF
END_IF

(* —— 段 9：故障/失能强制阀位全关（安全侧优先于段 8 联动） —— *)
IF (_eState <> E_DL_TbpState.eMonitor) THEN
    _bMakeup := FALSE;                                       // 非监测相：补气阀关 / Non-monitoring: make-up closed
    _bVent   := FALSE;                                       // 非监测相：排放阀关 / Non-monitoring: vent closed
    _fPct    := DL_TBP_PCT_MIN;                              // 非监测相：指令归零 / Non-monitoring: command zeroed
END_IF

(* —— 段 10：出口单点映射（名实双出口，R191） —— *)
fPrSelected   := _fSel;                                      // 可信压差出口 / Trusted pressure outlet
fPrDev        := _fDev;                                      // 双表偏差出口 / Deviation outlet
bMakeupValve  := _bMakeup;                                   // 补气阀位出口 / Make-up valve outlet
fValveCmdPct  := _fPct;                                      // 阀位指令出口（已限幅） / Command outlet, clamped
bVentValve    := _bVent;                                     // 排放阀位出口 / Vent valve outlet
bLowInterlock := _bLowLatch;                                 // 低压联锁出口 / Low interlock outlet
bSensorDev    := _bDevLatch;                                 // 双表偏离出口 / Deviation outlet
eState        := _eState;                                    // 相出口 / Phase outlet
eCause        := _eCause;                                    // 成因出口 / Cause outlet
bError        := _bFault OR _bDevLatch;                      // 故障标志（组态级或双表偏离） / Error flag

END_FUNCTION_BLOCK

(* ---- FB_DL_VacuumGaugeMux.st ---- *)
(*==============================================================================
 * 组件名称 (Component)  : FB_DL_VacuumGaugeMux
 * 所属子库 (Sublibrary) : DL_Device
 * 当前版本 (Version)    : 1.0.1
 * 组件分类 (Category)   : 功能块（FUNCTION_BLOCK）· 真空测量 · 双表量程选择与读数融合
 * 兼容性   (Platform)   : CODESYS 3.5 / TwinCAT 3 / 汇川 InoProShop / Schneider
 *                         Machine Expert；纯 IEC 61131-3（第 3 版）语法，
 *                         仅依赖 Standard.library（R_TRIG / LN / EXPT / ABS）
 * 功能描述 (Function)   : 皮拉尼（粗抽）与电容膜片（精抽）双真空计的量程选择、重叠区
 *                         交叉校验与读数融合。带切换迟滞防抖动、双表一致性判定、
 *                         不一致锁存与人工确认、以及按十倍程给出的偏差量化值。
 * 分层声明 (Layering)   : ① 本件只做「两表读数融合与一致性裁决」，不做采集调度、
 *                         不做线性化（皮拉尼的非线性修正由变送器或上位标定曲线承担）；
 *                         ② 不做腔体工艺联锁（联锁由工艺层消费融合后的单值压力）；
 *                         ③ 质量码复用设备层既有信号质量枚举，不另立质量枚举。
 * 不一致策略 (Disagree) : 不一致时**不死用任一表**：锁存不一致、置故障位、输出保持上次
 *                         值。理由：切换点附近两表差一个数量级时，无法判断是粗抽表污染
 *                         还是精抽表漂移，任选其一都可能把坏值送进工艺联锁。人工核后可
 *                         用确认沿清「不一致」标志，但故障锁存保留（诊断证据留存），
 *                         两条清除路径分离。
 * 融合规则 (Fusion)     : 重叠区内取电容膜片读数（精抽段比皮拉尼高一个数量级的精度，
 *                         属物理事实而非偏好）；重叠区外按当前选择表取原值。
 * 开源溯源 (Origin)     : 来源标签 namur-ne43 加 oscat-building。原创实现（参考 NAMUR
 *                         NE43「多段有效域 + 越域即诊断」的契约形态，以及 OSCAT Building
 *                         组「域外行为显式化」的写法）。仅借契约形态与参数域，切换迟滞、
 *                         十倍程交叉校验、融合规则、枚举、状态机与全部码位 100% 本库
 *                         独立设计，clean-room 实现，零代码行复制。OSCAT 为免费开源库，
 *                         此处按最严口径只借结构，不引其代码与注释。
 * 依赖     (Depends)    : E_DL_SignalQuality（设备层既有类型，本件只引用不声明）；
 *                         Standard.library: R_TRIG / LN / EXPT / ABS / LIMIT
 * 故障码表 (Error codes):
 *   16#0003_0153【信息级】重叠区宽度越界已钳到 0 至 3 个十倍程
 *   16#0003_0154【信息级】一致性容差越界已钳到 0.05 至 3 个十倍程
 *   16#0003_0155【信息级】仅单表可用，融合质量为不确定（不置故障位）
 *   16#0003_0313【故障级】切换点非正，量程划分无意义（锁存）
 *   16#0003_0314【故障级】双表不一致或双表均失效，输出保持（锁存）
 *   16#0003_0315【故障级】非法状态兜底（锁存，终端安全态）
 * 码位占用 (Slot)       : 信息级 0153 / 0154 / 0155；故障级 0313 / 0314 / 0315。
 *                         全部落在 R12 本件分配块内，无跨块借用、无段外哨兵值。
 * 拍序纪律 (Cycle order) :
 *   ① ePhase        ：段 6 状态机（唯一位移点），段 7 复位分支是唯一回退点
 *   ② fPressurePa   ：段 8 单点写出（成功拍写新值，其余拍回写保持值）
 *   ③ bDisagreeLatch：段 6 置位、段 7 由确认沿或复位沿清除，无第三处写入
 *   ④ uErrorId      ：段 9 单一优先级链，全拍只写一次
 * 验收向量 (Acceptance) :
 *   V1 重叠区外：皮拉尼 15、电容 12、切换点 10、重叠 1 个十倍程 → 下门限 3.162，
 *      15 高于上门限故不重叠，选皮拉尼，输出 15.0，不置不一致
 *   V2 不一致：皮拉尼 100、电容 1 → 偏差 2 个十倍程超过容差 0.5 → 锁不一致、
 *      故障位置位、码 0314、输出保持上次
 *   V3 重叠区一致：皮拉尼 6、电容 4 → 6 落在 3.162 到 10 之间，偏差 0.176 在容差内，
 *      取电容表 → 输出 4.0、采信表为电容、重叠标志为真、质量为良好
 *   V4 双表失效：两表有效位均假 → 故障位置位、码 0314、输出保持
 *   V5 迟滞：当前为皮拉尼、压力 8.0（高于下门限 3.162）→ 仍为皮拉尼，不切换
 * 偏离留档 (Deviation)  :
 *   ① 规格第 3.15 节正文写「重叠区内才交叉校验」，但验收向量 V2 的工况（100 与 1）
 *      并不落在重叠区，仍要求判不一致。本件按向量实现：只要两表都可用即做交叉校验
 *      （更保守），重叠区标志单独保留用于融合规则与画面提示。
 *   ② 质量码复用既有枚举，其成员语义按 NE43 四级设计，与本件的三档结论不是一一对应。
 *      本件在声明区定义三个映射基准量（良好、不确定、坏），使「本件结论到枚举」的
 *      对应关系只有一处，避免散落在各分支里出现多种写法。
 *   ③ 三相轮转（选择、校验、回选择）每拍推进一相，故同一路读数约两到三拍完成一次
 *      完整裁决；不采用单拍跑完两相，是为了让每个相位在画面上可观测。
 *   ④ 规格内部变量清单列有「双表均无效」标志量，本件在两处直接按条件进故障并置质量码，
 *      若保留该标志则只有写没有读（只置不销），故不声明，避免死状态量。
 * 修订历史 (Revision)   :
 *   2026-11-15  v1.0.0  首版落盘（R12 · 泳道 C · 双表真空计融合件）
 *   2026-11-15  v1.0.1  终审修复：融合发布增加「跨相失效保护」。选择相与本相相隔一拍，
 *                       若采信表在两拍之间掉线，原实现仍按该表原值（可能是 0 或负值）
 *                       写进 fPressurePa，与本件「不死用任一表」的契约相反；改为取值表
 *                       本拍不可用即不发布（bUpdateOut 取该表可用性），输出保持上次值，
 *                       下拍回选择相重新裁决
 *============================================================================*)

(*------------------------------------------------------------------------------
 * 枚举: E_DL_GaugeSel（采信表选择，归属本功能块并同文件发布）
 *       Active gauge selection owned by this block
 *-----------------------------------------------------------------------------*)
TYPE E_DL_GaugeSel :
(
    eNone        := 0,   // 未选：上电首拍或复位后，等待首次量程判定 / Not selected yet, waiting for the first decision
    ePirani      := 10,  // 皮拉尼：粗抽段，覆盖大气到十帕量级 / Pirani gauge covering the roughing range
    eCapacitance := 20   // 电容膜片：精抽段，覆盖十帕到十毫帕量级 / Capacitance gauge covering the fine range
);
END_TYPE

(*------------------------------------------------------------------------------
 * 枚举: E_DL_GaugePhase（本块相位，归属本功能块并同文件发布）
 *       Phase enumeration owned by this block
 *-----------------------------------------------------------------------------*)
TYPE E_DL_GaugePhase :
(
    eIdle          := 0,   // 待机：未使能或参数闸门未过，输出保持 / Idle, disabled or the gate has not passed
    eSelect        := 10,  // 选择：有效性判定与带迟滞的量程选择 / Selection with hysteresis
    eOverlapCheck  := 20,  // 交叉校验：十倍程偏差比较、融合与质量定级 / Cross check, fusion and quality grading
    eFault         := 99   // 故障：切换点非法、双表失效、不一致或非法状态 / Fault, needs a reset to leave
);
END_TYPE

FUNCTION_BLOCK FB_DL_VacuumGaugeMux
VAR_INPUT
    bEnable          : BOOL;                        // 使能，FALSE 时保持上次输出 [-] / Enable, the last output is held while FALSE
    bReset           : BOOL;                        // 复位故障与不一致锁存，上升沿有效 [-] / Rising edge clears the fault and the disagreement latch
    bAcknowledge     : BOOL;                        // 人工确认不一致，上升沿有效，不清故障锁存 [-] / Rising edge acknowledges a disagreement, the fault latch stays
    fPiraniPa        : REAL;                        // 皮拉尼读数 [帕]，有效域大于 1 纳帕 / Pirani reading in pascals, must exceed one nanopascal
    bPiraniValid     : BOOL;                        // 皮拉尼数据有效 [-] / Pirani reading valid flag
    fCapacitancePa   : REAL;                        // 电容膜片读数 [帕]，有效域大于 1 纳帕 / Capacitance gauge reading in pascals
    bCapacitanceValid: BOOL;                        // 电容膜片数据有效 [-] / Capacitance reading valid flag
    fSwitchPa        : REAL := 10.0;                // 切换点，皮拉尼量程上限 [帕]，域大于 0 / Switchover pressure, must exceed zero
    fOverlapDecades  : REAL := 1.0;                 // 重叠区宽度 [十倍程]，域 0 到 3 / Overlap width in decades, zero to three
    fAgreeTolDecades : REAL := 0.5;                 // 交叉校验允许偏差 [十倍程]，域 0.05 到 3 / Agreement tolerance in decades
END_VAR
VAR_OUTPUT
    fPressurePa      : REAL;                        // 融合后压力 [帕] / Fused pressure in pascals
    eActiveGauge     : E_DL_GaugeSel;               // 当前采信表 [-] / Active gauge
    bInOverlap       : BOOL;                        // 处于重叠区 [-] / Inside the overlap band
    bDisagree        : BOOL;                        // 双表不一致锁存 [-] / Disagreement latched
    fDeltaDecades    : REAL;                        // 两表偏差 [十倍程]，单表可用时为 0 / Deviation in decades, zero when only one gauge is usable
    eQuality         : E_DL_SignalQuality;          // 融合结果质量，复用既有枚举 [-] / Fused quality, reuses the existing enumeration
    bError           : BOOL;                        // 故障级锁存，仅 0313 0314 0315 置位 [-] / Latched fault, only fault level codes set it
    uErrorId         : UDINT;                       // 事件码，0 表示无事件 [代码] / Event code, zero means none
    eState           : E_DL_GaugePhase;             // 主状态机当前相位 [-] / Current phase of the main state machine
END_VAR
VAR
    fbTrigReset      : R_TRIG;                      // 复位沿检测，主周期无条件刷新 [-] / Reset edge detector, refreshed unconditionally
    fbTrigAck        : R_TRIG;                      // 确认沿检测，主周期无条件刷新 [-] / Acknowledge edge detector, refreshed unconditionally
    ePhase           : E_DL_GaugePhase := E_DL_GaugePhase.eIdle; // 内部相位，对外经 eState 输出 [-] / Internal phase exported as eState
    bInit            : BOOL := FALSE;               // 首扫标志，初值 FALSE，判据取非 [-] / First-scan flag initialised FALSE
    bFaultLatch      : BOOL;                        // 故障锁存，仅复位分支清除 [-] / Fault latch, cleared by the reset path only
    bDisagreeLatch   : BOOL;                        // 不一致锁存，确认沿或复位沿清除 [-] / Disagreement latch, cleared by the acknowledge or the reset edge
    uErrInt          : UDINT;                       // 故障级码寄存，锁存型 [代码] / Latched fault level code register
    uInfoCode        : UDINT;                       // 本拍信息级码，每拍重算 [代码] / Info level code recomputed every scan
    fHiSwitch        : REAL := 10.0;                // 切到电容的上门限 [帕] / Upper switch threshold
    fLoSwitch        : REAL := 3.162;               // 切回皮拉尼的下门限 [帕] / Lower switch threshold
    fOverUse         : REAL := 1.0;                 // 生效重叠宽度 [十倍程] / Effective overlap width
    fTolUse          : REAL := 0.5;                 // 生效交叉校验容差 [十倍程] / Effective agreement tolerance
    fLogPir          : REAL;                        // 皮拉尼十倍程 [十倍程] / Pirani log10 value
    fLogCap          : REAL;                        // 电容十倍程 [十倍程] / Capacitance log10 value
    fSelPa           : REAL;                        // 当前采信表读数 [帕] / Reading of the selected gauge
    fNew             : REAL;                        // 本次融合结果 [帕] / Fused result of this scan
    fLast            : REAL;                        // 上次成功输出的压力 [帕] / Last successfully published pressure
    eSel             : E_DL_GaugeSel := E_DL_GaugeSel.eNone; // 本次选择结果 [-] / Selected gauge of this scan
    bPirOk           : BOOL;                        // 皮拉尼可用（有效且大于下限且有限）[-] / Pirani usable flag
    bCapOk           : BOOL;                        // 电容可用 [-] / Capacitance usable flag
    bPirFin          : BOOL;                        // 皮拉尼读数有限 [-] / Pirani reading finite flag
    bCapFin          : BOOL;                        // 电容读数有限 [-] / Capacitance reading finite flag
    bUpdateOut       : BOOL;                        // 本拍有新的融合结果 [-] / A new fused result is available
    eQualGood        : E_DL_SignalQuality := E_DL_SignalQuality.eGood;        // 质量映射基准：良好（声明区取值，体内只与基准量比较）[-] / Quality mapping baseline, good
    eQualUncertain   : E_DL_SignalQuality := E_DL_SignalQuality.eUnderRange;  // 质量映射基准：不确定（借欠量程位表达「量测可信度下降」）[-] / Quality mapping baseline, uncertain
    eQualBad         : E_DL_SignalQuality := E_DL_SignalQuality.eWireBreakLow; // 质量映射基准：坏（借线路故障位表达「不可采信」）[-] / Quality mapping baseline, bad
END_VAR
VAR CONSTANT
    DL_LN10          : REAL := 2.302585093;         // 十的自然对数 [-] / Natural logarithm of ten
    DL_P_MIN         : REAL := 1.0E-9;              // 最小可接受压力 [帕]，防对数域零与负 / Minimum acceptable pressure preventing log of zero
    DL_P_MAX         : REAL := 1.0E9;               // 压力合理上限，超出视为非有限 [帕] / Pressure sanity limit
    DL_SWITCH_HYST   : REAL := 0.5;                 // 迟滞系数，重叠宽度的一半用于下门限 / Hysteresis factor, half of the overlap width
    DL_DEC_MIN       : REAL := 0.0;                 // 重叠宽度下限 [十倍程] / Lower overlap width
    DL_DEC_MAX       : REAL := 3.0;                 // 重叠宽度上限 [十倍程] / Upper overlap width
    DL_TOL_MIN       : REAL := 0.05;                // 容差下限 [十倍程] / Lower tolerance
    DL_TOL_MAX       : REAL := 3.0;                 // 容差上限 [十倍程] / Upper tolerance
    DL_ONE           : REAL := 1.0;                 // 实数一，防魔数 [无量纲] / Real one used instead of a magic number
END_VAR

(*------------------------------------------------------------------------------
 * 段 1｜输出确定性默认值（单拍标志与派生量每拍预清零，R25 第一律）
 *      Deterministic defaults first, derived flags pre-cleared every scan
 *-----------------------------------------------------------------------------*)
uInfoCode    := 16#0000_0000;                   // 信息级码每拍重算（Info code recomputed every scan）
bInOverlap   := FALSE;                          // 重叠标志预清零（Overlap flag pre-cleared）
fDeltaDecades := 0.0;                           // 偏差量预清零（Deviation pre-cleared）
bUpdateOut   := FALSE;                          // 融合更新标志预清零（Fused update flag pre-cleared）
bPirFin      := FALSE;                          // 皮拉尼有限标志预清零（Pirani finite flag pre-cleared）
bCapFin      := FALSE;                          // 电容有限标志预清零（Capacitance finite flag pre-cleared）

(*------------------------------------------------------------------------------
 * 段 2｜沿检测无条件刷新（红线：实例在 CASE 之外每拍必刷）
 *      Edge detection refreshed unconditionally outside the CASE
 *-----------------------------------------------------------------------------*)
fbTrigReset(CLK := bReset);
fbTrigAck(CLK := bAcknowledge);

(*------------------------------------------------------------------------------
 * 段 3｜首扫初始化（唯一合法范式：初值 FALSE，判据取非）
 *      First-scan initialisation following the single legal pattern
 *-----------------------------------------------------------------------------*)
IF NOT bInit THEN
    fLast          := 0.0;                      // 上次输出压力清零（Last pressure cleared）
    fNew           := 0.0;                      // 融合中间量清零（Fused temporary cleared）
    eSel           := E_DL_GaugeSel.eNone;      // 采信表置未选（Gauge selection reset）
    bFaultLatch    := FALSE;                    // 故障锁存清零（Fault latch cleared）
    bDisagreeLatch := FALSE;                    // 不一致锁存清零（Disagreement latch cleared）
    uErrInt        := 16#0000_0000;             // 故障码清零（Fault code cleared）
    fPressurePa    := 0.0;                      // 压力出口清零（Pressure outlet cleared）
    eActiveGauge   := E_DL_GaugeSel.eNone;      // 采信表出口置未选（Gauge outlet reset）
    eQuality       := eQualUncertain;           // 质量出口置不确定（Quality outlet set to uncertain）
    ePhase         := E_DL_GaugePhase.eIdle;    // 相位复位为待机（Phase reset to idle）
    bInit          := TRUE;                     // 首扫只做一次（First scan runs once）
END_IF

(*------------------------------------------------------------------------------
 * 段 4｜参数闸门（切换点非正属故障级；重叠宽度与容差越界属信息级，只钳位）
 *      Parameter gate, only the switchover pressure is fault level
 *-----------------------------------------------------------------------------*)
IF fSwitchPa <= DL_P_MIN THEN
    bFaultLatch := TRUE;                        // 切换点非法：锁故障（Illegal switchover pressure, latch a fault）
    uErrInt     := 16#0003_0313;                // 0313 切换点非正（Switchover pressure not positive）
    fHiSwitch   := DL_ONE;                      // 门限给安全值，避免本拍出现零除（Safe threshold avoids a division by zero）
    fLoSwitch   := DL_ONE;                      // 下门限同样给安全值（Lower threshold set to the safe value）
ELSE
    fHiSwitch := fSwitchPa;                     // 上门限即切换点（Upper threshold is the switchover pressure）
    IF fOverlapDecades < DL_DEC_MIN THEN
        fOverUse   := DL_DEC_MIN;               // 负宽度无意义：钳到 0（Negative width clamped to zero）
        uInfoCode  := 16#0003_0153;             // 0153 重叠宽度越界已钳位（Overlap width clamped）
    ELSIF fOverlapDecades > DL_DEC_MAX THEN
        fOverUse   := DL_DEC_MAX;               // 超上限钳位（Clamped to the upper bound）
        uInfoCode  := 16#0003_0153;             // 0153 重叠宽度越界已钳位（Overlap width clamped）
    ELSE
        fOverUse   := fOverlapDecades;          // 合法宽度直通（Valid width passed through）
    END_IF
    fLoSwitch := fSwitchPa / EXPT(10.0, fOverUse * DL_SWITCH_HYST); // 下门限按半宽十倍程折算（Lower threshold from half of the overlap width）
END_IF

IF fAgreeTolDecades < DL_TOL_MIN THEN
    fTolUse   := DL_TOL_MIN;                    // 容差下限钳位（Tolerance clamped to the lower bound）
    uInfoCode := 16#0003_0154;                  // 0154 容差越界已钳位（Tolerance clamped）
ELSIF fAgreeTolDecades > DL_TOL_MAX THEN
    fTolUse   := DL_TOL_MAX;                    // 容差上限钳位（Tolerance clamped to the upper bound）
    uInfoCode := 16#0003_0154;                  // 0154 容差越界已钳位（Tolerance clamped）
ELSE
    fTolUse   := fAgreeTolDecades;              // 合法容差直通（Valid tolerance passed through）
END_IF

(*------------------------------------------------------------------------------
 * 段 5｜有限性闸门与可用性判定（对数域前置拦截：零与负数在取对数前剔除）
 *      Finiteness gate and usability check, guarding the logarithm domain
 *-----------------------------------------------------------------------------*)
bPirFin := NOT ((fPiraniPa <> fPiraniPa) OR (ABS(fPiraniPa) > DL_P_MAX)); // 皮拉尼有限判定（Pirani finiteness test）
bCapFin := NOT ((fCapacitancePa <> fCapacitancePa) OR (ABS(fCapacitancePa) > DL_P_MAX)); // 电容有限判定（Capacitance finiteness test）
bPirOk  := bPiraniValid AND bPirFin AND (fPiraniPa >= DL_P_MIN);   // 三道闸：有效位、有限、大于下限（Three gates）
bCapOk  := bCapacitanceValid AND bCapFin AND (fCapacitancePa >= DL_P_MIN); // 三道闸：有效位、有限、大于下限（Three gates）

(*------------------------------------------------------------------------------
 * 段 6｜主状态机（枚举每个成员均有标签，末尾 ELSE 兜底到终端安全态）
 *      Main state machine, one label per member plus a trailing ELSE fallback
 *-----------------------------------------------------------------------------*)
CASE ePhase OF

    E_DL_GaugePhase.eIdle: // 待机：故障或未使能则停留，否则进入选择
        IF bFaultLatch THEN
            ePhase := E_DL_GaugePhase.eFault;   // 参数已锁故障：进故障态（Gate failed, enter the fault state）
        ELSIF bEnable THEN
            ePhase := E_DL_GaugePhase.eSelect;  // 进选择态（Enter the selection phase）
        END_IF

    E_DL_GaugePhase.eSelect: // 选择：先判双表失效，再按迟滞维持或切换
        IF (NOT bPirOk) AND (NOT bCapOk) THEN
            IF NOT bFaultLatch THEN
                bFaultLatch := TRUE;            // 锁故障，保留首出码（Latch the fault keeping the first code）
                uErrInt     := 16#0003_0314;    // 0314 双表失效（Both gauges failed）
            END_IF
            eQuality := eQualBad;               // 质量定为坏（Quality marked bad）
            ePhase   := E_DL_GaugePhase.eFault; // 进故障态（Enter the fault state）
        ELSE
            IF eSel = E_DL_GaugeSel.eNone THEN
                (* 首次选择：能进精抽段（读数不高于切换点）就先上电容表，否则用皮拉尼 *)
                IF bCapOk AND bPirOk THEN
                    IF fPiraniPa <= fHiSwitch THEN
                        eSel := E_DL_GaugeSel.eCapacitance; // 已在精抽段（Already in the fine range）
                    ELSE
                        eSel := E_DL_GaugeSel.ePirani;      // 仍在大气压侧（Still on the atmosphere side）
                    END_IF
                ELSIF bCapOk THEN
                    eSel := E_DL_GaugeSel.eCapacitance;     // 只有电容可用（Only the capacitance gauge is usable）
                ELSE
                    eSel := E_DL_GaugeSel.ePirani;          // 只有皮拉尼可用（Only the Pirani gauge is usable）
                END_IF
            END_IF
            IF eSel = E_DL_GaugeSel.ePirani THEN
                IF (NOT bPirOk) AND bCapOk THEN
                    eSel := E_DL_GaugeSel.eCapacitance; // 皮拉尼失效即切电容（Pirani lost, switch over at once）
                ELSIF bCapOk AND (fPiraniPa <= fLoSwitch) THEN
                    eSel := E_DL_GaugeSel.eCapacitance; // 降到下门限以下才切（Switch only below the lower threshold）
                END_IF
            ELSIF eSel = E_DL_GaugeSel.eCapacitance THEN
                IF (NOT bCapOk) AND bPirOk THEN
                    eSel := E_DL_GaugeSel.ePirani;      // 电容失效即切皮拉尼（Capacitance lost, switch back at once）
                ELSIF bPirOk AND (fCapacitancePa >= fHiSwitch) THEN
                    eSel := E_DL_GaugeSel.ePirani;      // 升到上门限以上才切（Switch only above the upper threshold）
                END_IF
            ELSE
                eSel := E_DL_GaugeSel.ePirani;          // 未选态残留兜底（Defensive fallback for the unselected state）
            END_IF
            ePhase := E_DL_GaugePhase.eOverlapCheck;    // 进交叉校验态（Enter the cross check phase）
        END_IF

    E_DL_GaugePhase.eOverlapCheck: // 交叉校验与融合
        IF eSel = E_DL_GaugeSel.eCapacitance THEN
            fSelPa := fCapacitancePa;               // 采信表读数取电容（Reading of the selected gauge）
        ELSE
            fSelPa := fPiraniPa;                    // 采信表读数取皮拉尼（Reading of the selected gauge）
        END_IF
        bInOverlap := (fSelPa >= fLoSwitch) AND (fSelPa <= fHiSwitch); // 重叠区判定（Overlap band test）
        fLogPir := 0.0;                             // 十倍程预清零（Log value pre-cleared）
        fLogCap := 0.0;                             // 十倍程预清零（Log value pre-cleared）
        IF bPirOk THEN
            fLogPir := LN(fPiraniPa) / DL_LN10;     // 取对数，前置闸门已排除零与负（Log guarded by the usability gate）
        END_IF
        IF bCapOk THEN
            fLogCap := LN(fCapacitancePa) / DL_LN10; // 取对数，前置闸门已排除零与负（Log guarded by the usability gate）
        END_IF
        IF bPirOk AND bCapOk THEN
            fDeltaDecades := ABS(fLogPir - fLogCap); // 两表偏差量化到十倍程（Deviation quantified in decades）
        END_IF
        IF (NOT bPirOk) AND (NOT bCapOk) THEN
            IF NOT bFaultLatch THEN
                bFaultLatch := TRUE;                // 锁故障（Latch the fault）
                uErrInt     := 16#0003_0314;        // 0314 双表失效（Both gauges failed）
            END_IF
            eQuality := eQualBad;                   // 质量定为坏（Quality marked bad）
            ePhase   := E_DL_GaugePhase.eFault;     // 进故障态（Enter the fault state）
        ELSIF bPirOk AND bCapOk AND (fDeltaDecades > fTolUse) THEN
            bDisagreeLatch := TRUE;                 // 锁不一致（Latch the disagreement）
            IF NOT bFaultLatch THEN
                bFaultLatch := TRUE;                // 锁故障（Latch the fault）
                uErrInt     := 16#0003_0314;        // 0314 双表不一致（Gauges disagree）
            END_IF
            eQuality := eQualBad;                   // 质量定为坏（Quality marked bad）
            ePhase   := E_DL_GaugePhase.eFault;     // 进故障态，输出保持（Enter the fault state, output held）
        ELSE
            IF bInOverlap AND bCapOk THEN
                fNew := fCapacitancePa;             // 重叠区取电容（融合取电容表） / Fusion takes the capacitance gauge in the overlap band
                bUpdateOut := TRUE;                 // 取值前已验可用，本拍有新结果 / The source was validated, publish it
            ELSE
                (* 重叠区外按选择表取原值：三个成员逐个给出取值口径，不留隐式分支 *)
                (* Outside the overlap band the selected gauge is used, one explicit label per member *)
                CASE eSel OF
                    E_DL_GaugeSel.eNone:
                        fNew := fPiraniPa;          // 未选态兜底取皮拉尼（Unselected fallback uses the Pirani gauge）
                    E_DL_GaugeSel.ePirani:
                        fNew := fPiraniPa;          // 选皮拉尼（The Pirani gauge is selected）
                    E_DL_GaugeSel.eCapacitance:
                        fNew := fCapacitancePa;     // 选电容膜片（The capacitance gauge is selected）
                    ELSE
                        fNew := fPiraniPa;          // 非法枚举值兜底（Illegal enumeration value fallback）
                END_CASE
                (* 跨相失效保护：选择相与本相相隔一拍，读数可能已掉线，取值表本拍不可用即不发布 *)
                (* Cross-phase guard: the selected gauge may have dropped out between the two phases *)
                IF eSel = E_DL_GaugeSel.eCapacitance THEN
                    bUpdateOut := bCapOk;           // 采信电容：本拍仍可用才发布 / Publish only while the capacitance gauge is usable
                ELSE
                    bUpdateOut := bPirOk;           // 采信皮拉尼：本拍仍可用才发布 / Publish only while the Pirani gauge is usable
                END_IF
            END_IF
            IF bPirOk AND bCapOk THEN
                eQuality := eQualGood;              // 双表可用且一致：良好（Both usable and consistent, good）
            ELSE
                eQuality := eQualUncertain;         // 单表可用：不确定（Single gauge, uncertain）
                uInfoCode := 16#0003_0155;          // 0155 单表可用（Single gauge usable）
            END_IF
            ePhase := E_DL_GaugePhase.eSelect;      // 回选择态，下拍重新判定（Back to selection）
        END_IF

    E_DL_GaugePhase.eFault: // 故障：输出保持，等复位沿（Fault, outputs held until the reset edge）
        eQuality := eQualBad;                       // 故障期质量定为坏（Quality marked bad during a fault）

    ELSE
        bFaultLatch := TRUE;                        // 非法状态兜底锁存（Illegal state latched）
        uErrInt     := 16#0003_0315;                // 0315 非法状态兜底（Illegal state fallback code）
        ePhase      := E_DL_GaugePhase.eFault;      // 进终端安全态（Enter the terminal safe state）
END_CASE

(*------------------------------------------------------------------------------
 * 段 7｜人工确认与复位（确认只清不一致标志，复位清故障锁存，两条路径分离）
 *      Acknowledge clears only the disagreement; reset clears the fault latch
 *-----------------------------------------------------------------------------*)
IF fbTrigAck.Q THEN
    bDisagreeLatch := FALSE;                    // 人工已核：清不一致（Acknowledged, clear the disagreement）
END_IF
IF fbTrigReset.Q THEN
    bDisagreeLatch := FALSE;                    // 复位清不一致（Reset clears the disagreement）
    bFaultLatch    := FALSE;                    // 复位清故障锁存（Reset clears the fault latch）
    uErrInt        := 16#0000_0000;             // 复位清故障码（Reset clears the fault code）
    eSel           := E_DL_GaugeSel.eNone;      // 选择表回未选，重新按读数判定（Selection reset to unselected）
    IF ePhase = E_DL_GaugePhase.eFault THEN
        ePhase := E_DL_GaugePhase.eIdle;        // 故障态复位回待机（Fault returns to idle）
    END_IF
END_IF

(*------------------------------------------------------------------------------
 * 段 8｜压力出口单点写出（成功拍写新值并刷新保持寄存器，其余拍回写保持值）
 *      Single write point of the pressure outlet with an explicit hold register
 *-----------------------------------------------------------------------------*)
IF bUpdateOut THEN
    fPressurePa := fNew;                        // 成功拍写出新值（Publish the new value）
    fLast       := fNew;                        // 刷新保持寄存器（Refresh the hold register）
ELSE
    fPressurePa := fLast;                       // 其余拍回写保持值，杜绝坏表值进联锁（Hold the last good value）
END_IF

(*------------------------------------------------------------------------------
 * 段 9｜码位定级与出口（单一优先级链，全拍只写一次 uErrorId）
 *      Single priority chain and outlet mapping
 *-----------------------------------------------------------------------------*)
eActiveGauge := eSel;                           // 采信表出口（Active gauge outlet）
bDisagree    := bDisagreeLatch;                 // 不一致出口（Disagreement outlet）
eState       := ePhase;                         // 相位出口（Phase outlet）
bError       := bFaultLatch;                    // 故障位只反映故障级锁存（Fault bit reflects the latch only）
IF bError THEN
    uErrorId := uErrInt;                        // 故障级码优先透出（Fault level code has priority）
ELSE
    uErrorId := uInfoCode;                      // 无故障透出本拍信息级码（Info code exposed otherwise）
END_IF
END_FUNCTION_BLOCK

(* ---- I_DL_AnalogSensor.st ---- *)
(*==============================================================================
 * 组件名称 (Component)  : I_DL_AnalogSensor
 * 所属子库 (Sublibrary) : DL_Device
 * 当前版本 (Version)    : 1.0.1
 * 兼容性   (Platform)   : CODESYS 3.5 / TwinCAT 3 / 汇川 InoProShop / Machine Expert
 *                         纯 IEC 61131-3（第3版）接口语法，零厂商方言
 * 分类     (Category)   : 设备抽象接口（Interface）+ 配套质量枚举（DUT）
 * 功能简述 (Function)   : 模拟量变送器标准抽象契约（NAMUR NE43 语义域）。
 *                         定义工程量当前值、信号质量分级、HH/H/L/LL 四级
 *                         报警位与故障码的只读属性组，供温控区（如
 *                         FB_DL_HeatCoolZone）等上层工艺块做依赖注入；
 *                         原始信号采集、标定与诊断由实现块
 *                         （如 FB_DL_AnalogTransmitter）完成。
 * 开源溯源 (Origin)     : 来源标签 namur-ne43（RAW_NOTES_R5 S-5：NAMUR NE43
 *                         信号电平域为公开推荐实践，多来源交叉印证——
 *                         有效测量域 3.8~20.5 mA、故障域 <3.6 / >21 mA、
 *                         0 mA 回路断线、超量程标记而非剔除；仅借鉴公开
 *                         标准语义，接口命名、质量分级枚举按本库红线独立
 *                         设计，clean-room 未复制任何源码行）。
 * 红线自检 (Redline)    : R1 零全局变量表/外部变量引用 ✓｜R2 零物理 IO 地址 ✓
 *                         R3 纯 IEC 61131-3 ✓｜R5 全成员中英双语同行注释 ✓
 *                         R18 接口以 END_INTERFACE 成对终结 ✓
 * 归属说明 (Ownership)  : 本文件同时承载 E_DL_SignalQuality 枚举定义，
 *                         该枚举归属接口 I_DL_AnalogSensor，与其同文件发布。
 * 修订历史 (Revision)   :
 *   2026-11-15  v1.0.0  首版入库（R5 轮 · DL_Device 开库）
 *   2026-11-15  v1.0.1  R11 修复：枚举成员分隔符笔误，eWireBreakLow / eWireBreakHigh 两行误写单冒号 `:`（IEC 61131-3 枚举成员赋值须用 `:=`），三平台编译阻断已消除，数值与语义不变。
 *                       R11 fix: enum member separator erratum, `:` -> `:=` on two members.
 *============================================================================*)

(*-----------------------------------------------------------------------------
 * 枚举: E_DL_SignalQuality（归属接口 I_DL_AnalogSensor，与其同文件）
 * 含义: NAMUR NE43 信号质量分级。数值步长 10 留空位，便于后续插态；
 *       断线/开路三个诊断态取 30/40/50 依严重度递增排序。
 *----------------------------------------------------------------------------*)
TYPE E_DL_SignalQuality :
(
    eGood         := 0,    // 信号良好：原始值位于有效测量域内 / Signal good, raw value inside valid measurement span
    eUnderRange   := 10,   // 欠量程：原始值低于量程下限但在故障门限之上（如 3.8~4.0 mA 段）/ Under-range, raw below span low but above fault threshold
    eOverRange    := 20,   // 超量程：原始值高于量程上限但在故障门限之下（如 20.0~20.5 mA 段）/ Over-range, raw above span high but below fault threshold
    eWireBreakLow := 30,   // 低侧断线：原始值低于故障下门限（如 <3.6 mA，按配置方向判定）/ Wire break low side, raw below low fault threshold per configured direction
    eWireBreakHigh := 40,  // 高侧断线：原始值高于故障上门限（如 >21 mA，按配置方向判定）/ Wire break high side, raw above high fault threshold per configured direction
    eOpenLoop     := 50    // 回路开路：原始值接近 0 域（0 mA/0 V），变送器失电或回路断开 / Open loop, raw near zero domain, loop broken or transmitter unpowered
) USINT;
END_TYPE

(*-----------------------------------------------------------------------------
 * 接口: I_DL_AnalogSensor
 * 契约结构: 属性（PROPERTY GET）单段式，方法总数 0 个，远低于 ≤6 红线；
 *           纯只读数据契约——诊断与标定逻辑全部驻留实现块内部。
 * 边界防错: fValue 输出承诺经非有限值防御（输入为非数时保持末次有效值），
 *           调用方无需再做空值判护；故障态下 fValue 保持末次有效工程量
 *           并由 eQuality 与 uErrorId 显式标注，杜绝把故障电流当过程值。
 *----------------------------------------------------------------------------*)
INTERFACE I_DL_AnalogSensor

// ---- 属性段（全部只读 GET）------------------------------------------------

PROPERTY fValue    : REAL              // 工程量当前值（Current engineering value），单位由调用方标定组态约定，故障态保持末次有效值 / Current value, unit per caller scaling config, holds last good value in fault
PROPERTY eQuality  : E_DL_SignalQuality // 信号质量分级（Signal quality grade），NE43 四段诊断结果 / NE43 diagnostic grade
PROPERTY bAlarmHH  : BOOL              // 上上限报警（High-high alarm），TRUE=工程量越上上限门限 / TRUE = value above high-high limit
PROPERTY bAlarmH   : BOOL              // 上限报警（High alarm），TRUE=工程量越上限门限 / TRUE = value above high limit
PROPERTY bAlarmL   : BOOL              // 下限报警（Low alarm），TRUE=工程量越下限门限 / TRUE = value below low limit
PROPERTY bAlarmLL  : BOOL              // 下下限报警（Low-low alarm），TRUE=工程量越下下限门限 / TRUE = value below low-low limit
PROPERTY uErrorId  : UDINT             // 末次故障码（Last error code），0=无故障，段位 16#0003_xxxx / Last error code, 0 = none, family 16#0003_xxxx

END_INTERFACE
